(* CODESYS project i_hmi.library
   DefaultNamespace: KOSTAL.AF2024.HMI.I_Hmi
   DocFormat: reStructuredText
   Description: Base for HMI Interfaces in UTF16
   Author: Frank Dümpelmann
   Title: KOSTAL.AF2024.HMI.I_Hmi
   Version: 1.0.0.0
   Company: KOSTAL GmbH & Co.KG
   Placeholder: KOSTAL.AF2024.HMI.I_Hmi

Project tree, tasks and I/O mapping:
  libraries: KOSTAL.AF2024.Core.functionResponse, 1.0.0.0 (KOSTAL GmbH & Co.KG); KOSTAL.AF2024.Core.MainControl, 1.0.0.0 (KOSTAL GmbH & Co.KG); KOSTAL.AF2024.Core.Process, 1.0.0.0 (KOSTAL GmbH & Co.KG); KOSTAL.AF2024.Core.Settings, 1.0.0.0 (KOSTAL GmbH & Co.KG); KOSTAL.AF2024.Core.System, 1.0.0.0 (KOSTAL GmbH & Co.KG); KOSTAL.AF2024.HMI.Controls, 1.0.0.0 (KOSTAL GmbH & Co.KG)
  Aliases/
    data type T_ARTICLENAME
    data type T_BUTTON_TEXT
    data type T_F_BUTTON_TEXT
    data type T_LANGUAGENAME
    data type T_PAGE_TEXT
  DUT/
    Fn_Button/
      interface _I_T_Fn_Button: Button, clear_controls
      interface _I_T_Fn_Button_CopyFrom: CopyFrom
      interface _I_T_Fn_Button_Owner: Button_Owner, clear, clear_signals, CopyFrom
      interface _I_T_Fn_Button_RO: Button_RO, CopyTo
      data type _T_F_ButtonRange
      function block _T_Fn_Button [ST]: Button, Button_Owner, Button_RO, clear, clear_controls, clear_signals, CopyFrom, CopyTo
    Message/
      interface _I_T_Message: clear, Content, State
      interface _I_T_Message_CopyFrom: CopyFrom
      interface _I_T_Message_Owner: CopyFrom
      interface _I_T_Message_RO: Content, CopyTo, State
      function block _T_Message [ST]: clear, Content, CopyFrom, CopyTo, State
    data type E_STATE
    data type E_UserLevel
  MainControl/
    function block FB_MainControl [ST]: Button_Article_Owner, Button_Auto_Owner, Button_Door_Owner, Button_Manual_Owner, Button_OnOff_Owner, Button_Parameters_Owner, Button_Run_Owner, Button_RunEmpty_Owner, Button_Article_RO, Button_Auto_RO, Button_Door_RO, Button_Manual_RO, Button_OnOff_RO, Button_Parameters_RO, Button_Run_RO, Button_RunEmpty_RO, Button_Article, Button_Auto, Button_Door, Button_Manual, Button_OnOff, Button_Parameters, Button_RunEmpty, Button_RunStop, clear, Language, linkMainControl, Name, statusDoor_close, statusDoor_open, statusDoor_safe, UserLevel, Version_PLC
    interface I_MainControl: Button_Article, Button_Auto, Button_Door, Button_Manual, Button_OnOff, Button_Parameters, Button_RunEmpty, Button_RunStop, Language, linkMainControl, Name, statusDoor_close, statusDoor_open, statusDoor_safe, UserLevel, Version_PLC
    interface I_MainControl_Owner: Button_Article_Owner, Button_Auto_Owner, Button_Door_Owner, Button_Manual_Owner, Button_OnOff_Owner, Button_Parameters_Owner, Button_Run_Owner, Button_RunEmpty_Owner, Language, clear
    interface I_MainControl_RO: Button_Article_RO, Button_Auto_RO, Button_Door_RO, Button_Manual_RO, Button_OnOff_RO, Button_Parameters_RO, Button_Run_RO, Button_RunEmpty_RO, Language, Name, statusDoor_close, statusDoor_open, statusDoor_safe, UserLevel, Version_PLC
  Page/
    Page_Listing/
      _Buttons/
        interface _I_T_Listing_Buttons: Button_Left, Button_Right, clear_controls
        interface _I_T_Listing_Buttons_CopyFrom: CopyFrom
        interface _I_T_Listing_Buttons_Owner: Button_Left_Owner, Button_Right_Owner, clear, clear_signals, CopyFrom
        interface _I_T_Listing_Buttons_RO: Button_Right_RO, Button_RO, CopyTo
        function block _T_Listing_Buttons [ST]: Button_Left, Button_Left_Owner, Button_Right, Button_Right_Owner, Button_Right_RO, Button_RO, clear, clear_controls, clear_signals, CopyFrom, CopyTo
      _Messages/
        interface _I_T_Listing_Messages: clear, Message
        interface _I_T_Listing_Messages_CopyFrom: CopyFrom
        interface _I_T_Listing_Messages_Owner: CopyFrom, Message_Owner
        interface _I_T_Listing_Messages_RO: CopyTo, Message_RO
        function block _T_Listing_Messages [ST]: clear, CopyFrom, CopyTo, Message, Message_Owner, Message_RO
      Listing/
        function block FB_Page_Listing [ST]: Activate, Buttons, Buttons_Owner, Buttons_RO, clear, clear_buttons, clear_controls, clear_messages, clear_signals, Messages, Messages_Owner, Messages_RO
        interface I_Page_Listing: Activate, Buttons, clear_controls, clear_messages, Messages
        interface I_Page_Listing_Owner: Buttons_Owner, clear, clear_buttons, clear_signals, Messages_Owner
        interface I_Page_Listing_RO: Activate, Buttons_RO, Messages_RO
    Page_PDEF/
      _Button/
        interface _I_T_PDEF_Button_Member: State
        interface _I_T_PDEF_Button_Owner: State
        interface _I_T_PDEF_Button_RO: State
        function block _T_PDEF_Button [ST]: clear, clear_control, CopyFrom, State
      _Buttons/
        interface _I_T_PDEF_Buttons_CopyFrom: CopyFrom
        interface _I_T_PDEF_Buttons_Member: Button_Member, clear_controls
        interface _I_T_PDEF_Buttons_Owner: Button_Owner, clear, clear_signals, CopyFrom
        interface _I_T_PDEF_Buttons_RO: Button, CopyTo
        function block _T_PDEF_Buttons [ST]: Button, Button_Member, Button_Owner, clear, clear_controls, clear_signals, CopyFrom, CopyTo
      _Messages/
        interface _I_T_PDEF_Messages_CopyFrom: CopyFrom
        interface _I_T_PDEF_Messages_Member: clear, CopyFrom, Message
        interface _I_T_PDEF_Messages_Owner: Message_Owner
        interface _I_T_PDEF_Messages_RO: CopyTo, Message_RO
        function block _T_PDEF_Messages [ST]: clear, CopyFrom, CopyTo, Message, Message_Owner, Message_RO
      PDEF/
        function block FB_Page_PDEF [ST]: Buttons, Confirm, Message, Messages, Buttons_Owner, Confirm_Owner, Message_Owner, Messages_Owner, Buttons_RO, Confirm_RO, Message_RO, Messages_RO, Activate, clear, Name
        interface I_Page_PDEF: Buttons, Confirm, Message, Messages, Buttons_RO, Confirm_RO, Message_RO, Messages_RO, Activate, Name
        interface I_Page_PDEF_Owner: Buttons, Confirm, Message, Messages, Buttons_Owner, Confirm_Owner, Message_Owner, Messages_Owner, Buttons_RO, Confirm_RO, Message_RO, Messages_RO, Activate, clear, Name
        interface I_Page_PDEF_RO: Activate, Buttons_RO, Confirm_RO, Message_RO, Messages_RO, Name
    Page_Station/
      function block FB_Page_Station [ST]: Button_Enter, Button_Escape, Button_Minus, Button_OnOff, Button_Plus, Buttons_Custom, clear_controls, Name, Status, Text, Button_Enter_Owner, Button_Escape_Owner, Button_Minus_Owner, Button_OnOff_Owner, Button_Plus_Owner, Buttons_Custom_Owner, clear, clear_button, clear_signals, Status_Owner, Text_Owner, Button_Enter_RO, Button_Escape_RO, Button_Minus_RO, Button_OnOff_RO, Button_Plus_RO, Buttons_Custom_RO, Name_RO, Status_RO, Text_RO
      interface I_Page_Station: Button_Enter, Button_Escape, Button_Minus, Button_OnOff, Button_Plus, Buttons_Custom, clear_controls, Name, Status, Text
      interface I_Page_Station_Owner: Button_Enter_Owner, Button_Escape_Owner, Button_Minus_Owner, Button_OnOff_Owner, Button_Plus_Owner, Buttons_Custom_Owner, clear, clear_button, clear_signals, Status_Owner, Text_Owner
      interface I_Page_Station_RO: Button_Enter_RO, Button_Escape_RO, Button_Minus_RO, Button_OnOff_RO, Button_Plus_RO, Buttons_Custom_RO, Name, Status_RO, Text_RO
    Page_XYZ/
      _Buttons/
        interface _I_T_XYZ_Buttons: Button, clear_controls
        interface _I_T_XYZ_Buttons_CopyFrom: CopyFrom
        interface _I_T_XYZ_Buttons_Owner: Button_Owner, clear, clear_signals, CopyFrom
        interface _I_T_XYZ_Buttons_RO: Button_RO, CopyTo
        function block _T_XYZ_Buttons [ST]: Button, Button_Owner, Button_RO, clear, clear_controls, clear_signals, CopyFrom, CopyTo
      function block FB_page_XYZ [ST]: Button_Backward, Button_Down, Button_Forward, Button_Left, Button_Minus, Button_Plus, Button_Right, Button_Up, Buttons_Custom, clear_controls, SetText, Button_Backward_Owner, Button_Down_Owner, Button_Forward_Owner, Button_Left_Owner, Button_Minus_Owner, Button_Plus_Owner, Button_Right_Owner, Button_Up_Owner, Buttons_Custom_Owner, Button_Backward_RO, Button_Down_RO, Button_Forward_RO, Button_Left_RO, Button_Minus_RO, Button_Plus_RO, Button_Right_RO, Button_Up_RO, Buttons_Custom_RO, GetText, Activate, clear, clear_signals
      interface I_page_XYZ: Activate, Button_Backward, Button_Down, Button_Forward, Button_Left, Button_Minus, Button_Plus, Button_Right, Button_Up, clear_controls, SetText
      interface I_page_XYZ_Owner: Button_Backward_Owner, Button_Down_Owner, Button_Forward_Owner, Button_Left_Owner, Button_Minus_Owner, Button_Plus_Owner, Button_Right_Owner, Button_Up_Owner, clear, clear_signals
      interface I_page_XYZ_RO: Activate, Button_Backward_RO, Button_Down_RO, Button_Forward_RO, Button_Left_RO, Button_Minus_RO, Button_Plus_RO, Button_Right_RO, Button_Up_RO, GetText
  Project Information/
    function F_GetCompany [ST]
    function F_GetTitle [ST]
    function F_GetVersion [ST]
  Version/
    global variables Global_Version
  global variables GVL_CONSTANT
*)

// Aliases/T_ARTICLENAME
TYPE T_ARTICLENAME : STRING(40)
; END_TYPE

// Aliases/T_BUTTON_TEXT
TYPE T_BUTTON_TEXT : WSTRING(15)
; END_TYPE

// Aliases/T_F_BUTTON_TEXT
TYPE T_F_BUTTON_TEXT : WSTRING(10)
; END_TYPE

// Aliases/T_LANGUAGENAME
TYPE T_LANGUAGENAME : STRING(40)
; END_TYPE

// Aliases/T_PAGE_TEXT
TYPE T_PAGE_TEXT : WSTRING(255)
; END_TYPE

// DUT/Fn_Button/_T_F_ButtonRange
(*
Description
===========
| Limited data type for the index of an F-Button
*)
TYPE _T_F_ButtonRange : INT(1..8); END_TYPE

// DUT/E_STATE
(*
Description
===========
| Data type to describe a message state
*)
{attribute 'qualified_only'}
{attribute 'strict'}
TYPE E_STATE :
	(
		NONE						:=0, 
		PASS						:=1, 
		FAIL						:=2, 
		ATTENTION				:=3, 
		ERROR						:=4, 
		COMMON_REQUEST	:=5
	);
END_TYPE

// DUT/E_UserLevel
{attribute 'qualified_only'}
{attribute 'strict'}
TYPE E_UserLevel :
(
	operator := 0,
	service := 1,
	quality := 2
);
END_TYPE

// Version/Global_Version
{attribute 'TcGenerated'}
{attribute 'no-analysis'}
{attribute 'linkalways'}
// This function has been automatically generated from the project information.
VAR_GLOBAL CONSTANT
	{attribute 'const_non_replaced'}
	stLibVersion_KOSTAL_AF2024_HMI_I_Hmi : ST_LibVersion := (iMajor := 1, iMinor := 0, iBuild := 0, iRevision := 0, nFlags := 0, sVersion := '1.0.0.0');
END_VAR

// GVL_CONSTANT
{attribute 'qualified_only'}
VAR_GLOBAL CONSTANT

	MAX_FN_BUTTON	: INT:= 7;	//INT:= 7 	Maximum number of F-buttons (F8 is intern used as Help Page access)

	MAX_LISTING_LINE	: INT:= 10;	//INT:= 10	Maximum number of lines on listing page
	
	MAX_PDEF_BUTTONS	: INT:= 12;	//INT:= 12	Maximum number of FDEF buttons
	MAX_PDEF_MESSAGES	: INT:= 9;	//INT:= 9	Maximum number of FDEF messages

	MAX_XYZ_LINE	: INT:= 4;
	MAX_XYZ_BUTTON		: INT:= 4;	//INT:= 4	Maximum number of cusom Buttons on XYZ page
END_VAR

// DUT/Fn_Button/_I_T_Fn_Button
INTERFACE _I_T_Fn_Button EXTENDS _I_T_Fn_Button_RO

METHOD PUBLIC Button : KOSTAL_AF2024_HMI_Controls.I_T_Button_controlled
VAR_INPUT
	Number	: INT;
END_VAR
END_METHOD

METHOD PUBLIC clear_controls
END_METHOD

END_INTERFACE

// DUT/Fn_Button/_I_T_Fn_Button_RO
INTERFACE _I_T_Fn_Button_RO EXTENDS KOSTAL_AF2024_Core_System.I_Interface

METHOD PUBLIC Button_RO : KOSTAL_AF2024_HMI_Controls.I_T_Button_controlled
VAR_INPUT
	Number	: _T_F_ButtonRange;
END_VAR
END_METHOD

METHOD PUBLIC CopyTo
VAR_INPUT
	IN	: _I_T_Fn_Button_CopyFrom;
END_VAR
END_METHOD

END_INTERFACE

// DUT/Fn_Button/_I_T_Fn_Button_CopyFrom
INTERFACE _I_T_Fn_Button_CopyFrom EXTENDS KOSTAL_AF2024_Core_System.I_Interface

METHOD PUBLIC CopyFrom
VAR_INPUT
	IN	: _I_T_Fn_Button_RO;
END_VAR
END_METHOD

END_INTERFACE

// DUT/Fn_Button/_I_T_Fn_Button_Owner
INTERFACE _I_T_Fn_Button_Owner EXTENDS _I_T_Fn_Button

METHOD PUBLIC Button_Owner : KOSTAL_AF2024_HMI_Controls.I_T_Button_controlled_Owner
VAR_INPUT
	Number	: _T_F_ButtonRange;
END_VAR
END_METHOD

METHOD PUBLIC clear
END_METHOD

METHOD PUBLIC clear_signals
END_METHOD

METHOD PUBLIC CopyFrom
VAR_INPUT
	IN	: _I_T_Fn_Button_RO;
END_VAR
END_METHOD

END_INTERFACE

// DUT/Fn_Button/_T_Fn_Button
(*

:Author: Frank Dümpelmann <f.duempelmann@kostal.com>, Martin Hundt <m.hundt@kostal.com>
:Date: 2018-11-20

Function
========
| Data structure representing an array of buttons (FB_ControlledButton)
| Function to clear all content or signals only
*)

FUNCTION_BLOCK PUBLIC _T_Fn_Button IMPLEMENTS _I_T_Fn_Button_RO, _I_T_Fn_Button_Owner, _I_T_Fn_Button, _I_T_Fn_Button_CopyFrom

VAR
	_F		: ARRAY[1..GVL_CONSTANT.MAX_FN_BUTTON] OF KOSTAL_AF2024_HMI_Controls.T_Button_controlled;	//ARRAY[1..GVL_CONSTANT.MAX_FN_BUTTON] OF KOSTAL_TC3_Controls_button.FB_Button_controlled
	_Dummy	: KOSTAL_AF2024_HMI_Controls.T_Button_controlled;
END_VAR

METHOD PUBLIC Button : KOSTAL_AF2024_HMI_Controls.I_T_Button_controlled
VAR_INPUT
	Number	: INT;
END_VAR

IF (Number < 1) OR (Number > GVL_CONSTANT.MAX_FN_BUTTON) THEN	Button:= _Dummy;	RETURN;	END_IF

Button:= _F[Number];
END_METHOD

METHOD PUBLIC Button_Owner : KOSTAL_AF2024_HMI_Controls.I_T_Button_controlled_Owner
VAR_INPUT
	Number	: _T_F_ButtonRange;
END_VAR

IF (Number < 1) OR (Number > 8) THEN	Button_Owner:= _Dummy;	RETURN;	END_IF

Button_Owner:= _F[Number];
END_METHOD

METHOD PUBLIC Button_RO : KOSTAL_AF2024_HMI_Controls.I_T_Button_controlled
VAR_INPUT
	Number	: _T_F_ButtonRange;
END_VAR

IF (Number < 1) OR (Number > 8) THEN	Button_RO:= _Dummy;	RETURN;	END_IF

Button_RO:= _F[Number];
END_METHOD

METHOD PUBLIC clear


VAR
	_index: INT;	//INT
END_VAR

FOR _index:= 1 TO GVL_CONSTANT.MAX_FN_BUTTON DO
	_F[_index].clear();
END_FOR
END_METHOD

METHOD PUBLIC clear_controls

VAR
	_index: INT;	//INT
END_VAR

FOR _index:= 1 TO GVL_CONSTANT.MAX_FN_BUTTON DO
	_F[_index].clear_control();
END_FOR
END_METHOD

METHOD PUBLIC clear_signals

VAR
	_index: INT;	//INT
END_VAR

FOR _index:= 1 TO GVL_CONSTANT.MAX_FN_BUTTON DO
	_F[_index].clear_signals();
END_FOR
END_METHOD

METHOD PUBLIC CopyFrom
VAR_INPUT
	IN	: _I_T_Fn_Button_RO;
END_VAR

VAR
	_i: INT;
END_VAR

IF IN = 0 THEN RETURN;	END_IF

FOR _i:= 1 TO GVL_CONSTANT.MAX_FN_BUTTON DO
	_F[_i].CopyFrom(IN.Button_RO(_i));
END_FOR
END_METHOD

METHOD PUBLIC CopyTo
VAR_INPUT
	IN	: _I_T_Fn_Button_CopyFrom;
END_VAR

IF IN = 0 THEN RETURN;	END_IF

IN.CopyFrom(THIS^);
END_METHOD

END_FUNCTION_BLOCK

// DUT/Message/_I_T_Message
INTERFACE _I_T_Message EXTENDS _I_T_Message_RO

METHOD PUBLIC clear
VAR_INPUT
END_VAR
END_METHOD

PROPERTY PUBLIC Content : KOSTAL_AF2024_Core_Settings.T_MaxString
SET
END_SET
END_PROPERTY

PROPERTY PUBLIC State : E_STATE
SET
END_SET
END_PROPERTY

END_INTERFACE

// DUT/Message/_I_T_Message_RO
INTERFACE _I_T_Message_RO EXTENDS KOSTAL_AF2024_Core_System.I_Interface

PROPERTY PUBLIC Content : KOSTAL_AF2024_Core_Settings.T_MaxString
GET
END_GET
END_PROPERTY

METHOD PUBLIC CopyTo
VAR_INPUT
	IN	: _I_T_Message_CopyFrom;
END_VAR
END_METHOD

PROPERTY PUBLIC State : E_STATE
GET
END_GET
END_PROPERTY

END_INTERFACE

// DUT/Message/_I_T_Message_CopyFrom
INTERFACE _I_T_Message_CopyFrom EXTENDS KOSTAL_AF2024_Core_System.I_Interface

METHOD PUBLIC CopyFrom
VAR_INPUT
	IN	: _I_T_Message_RO;
END_VAR
END_METHOD

END_INTERFACE

// DUT/Message/_I_T_Message_Owner
INTERFACE _I_T_Message_Owner EXTENDS _I_T_Message

METHOD PUBLIC CopyFrom
VAR_INPUT
	IN	: _I_T_Message_RO;
END_VAR
END_METHOD

END_INTERFACE

// DUT/Message/_T_Message
(*

:Author: Frank Dümpelmann <f.duempelmann@kostal.com>, Martin Hundt <m.hundt@kostal.com>
:Date: 2018-11-20

Function
========
Data type representing a message with content (text) and state (error, pass,fail,...)

*)

FUNCTION_BLOCK PUBLIC _T_Message IMPLEMENTS _I_T_Message_RO, _I_T_Message_Owner, _I_T_Message, _I_T_Message_CopyFrom

VAR
	_Content	: KOSTAL_AF2024_Core_Settings.T_MaxString;
	_State		: E_STATE;
END_VAR

METHOD PUBLIC clear
VAR_INPUT
END_VAR

_Content:= "";
_State:= E_STATE.NONE;
END_METHOD

PROPERTY PUBLIC Content : KOSTAL_AF2024_Core_Settings.T_MaxString
GET

Content:= _Content;
END_GET
SET

_Content:= Content;
END_SET
END_PROPERTY

METHOD PUBLIC CopyFrom
VAR_INPUT
	IN	: _I_T_Message_RO;
END_VAR

IF IN = 0 THEN RETURN;	END_IF

_Content	:= IN.Content;
_State		:= IN.State;
END_METHOD

METHOD PUBLIC CopyTo
VAR_INPUT
	IN	: _I_T_Message_CopyFrom;
END_VAR

IF IN = 0 THEN RETURN;	END_IF

IN.CopyFrom(THIS^);
END_METHOD

PROPERTY PUBLIC State : E_STATE
GET

State:= _State;
END_GET
SET

_State:= State;
END_SET
END_PROPERTY

END_FUNCTION_BLOCK

// MainControl/FB_MainControl
(*

:Author: Frank Dümpelmann <f.duempelmann@kostal.com>, Martin Hundt <m.hundt@kostal.com>
:Date: 2020-02-20

Function
========
| Base class to implement a machine's main control

Methods and Properties
======================
| see documentation

*)
FUNCTION_BLOCK PUBLIC FB_MainControl IMPLEMENTS I_MainControl_RO, I_MainControl_Owner, I_MainControl

VAR
	_Name		: KOSTAL_AF2024_Core_Settings.T_MaxString;

	_OnOff		: KOSTAL_AF2024_HMI_Controls.T_Button_controlled;
	_RunStop	: KOSTAL_AF2024_HMI_Controls.T_Button_controlled;
	_RunEmpty	: KOSTAL_AF2024_HMI_Controls.T_Button_controlled;
                                             
	_Manual		: KOSTAL_AF2024_HMI_Controls.T_Button_controlled;
	_Auto		: KOSTAL_AF2024_HMI_Controls.T_Button_controlled;
	_Parameters		: KOSTAL_AF2024_HMI_Controls.T_Button_controlled;
	_Door		: KOSTAL_AF2024_HMI_Controls.T_Button_controlled;
	_Article	: KOSTAL_AF2024_HMI_Controls.T_Button_controlled;

	_statusDoor_close	: BOOL;	
	_statusDoor_open	: BOOL;	
	_statusDoor_safe	: BOOL;	
	
	_mainControl	: KOSTAL_AF2024_Core_MainControl.I_MainControl;

	
	_userLevel		: E_UserLevel;
	_language			: STRING;
	_version_PLC	: STRING;


END_VAR

(*
Description
===========
| Article button
*)
PROPERTY PUBLIC Button_Article_Owner : KOSTAL_AF2024_HMI_Controls.I_T_Button_controlled_Owner
GET

Button_Article_Owner := _Article;
END_GET
END_PROPERTY

(*
Description
===========
| Automatic button
*)
PROPERTY PUBLIC Button_Auto_Owner : KOSTAL_AF2024_HMI_Controls.I_T_Button_controlled_Owner
GET

Button_Auto_Owner := _Auto;
END_GET
END_PROPERTY

(*
Description
===========
| Door button
*)
PROPERTY PUBLIC Button_Door_Owner : KOSTAL_AF2024_HMI_Controls.I_T_Button_controlled_Owner
GET

Button_Door_Owner := _Door;
END_GET
END_PROPERTY

(*
Description
===========
| Manual button
*)
PROPERTY PUBLIC Button_Manual_Owner : KOSTAL_AF2024_HMI_Controls.I_T_Button_controlled_Owner
GET

Button_Manual_Owner := _Manual;
END_GET
END_PROPERTY

(*
Description
===========
| On/off button
*)
PROPERTY PUBLIC Button_OnOff_Owner : KOSTAL_AF2024_HMI_Controls.I_T_Button_controlled_Owner
GET

Button_OnOff_Owner := _OnOff;
END_GET
END_PROPERTY

(*
Description
===========
| Parameters button
*)
PROPERTY PUBLIC Button_Parameters_Owner : KOSTAL_AF2024_HMI_Controls.I_T_Button_controlled_Owner
GET

Button_Parameters_Owner := _Parameters;
END_GET
END_PROPERTY

(*
Description
===========
| Run button
*)

PROPERTY PUBLIC Button_Run_Owner : KOSTAL_AF2024_HMI_Controls.I_T_Button_controlled_Owner
GET

Button_Run_Owner := _RunStop;
END_GET
END_PROPERTY

(*
Description
===========
| Work empty button
*)
PROPERTY PUBLIC Button_RunEmpty_Owner : KOSTAL_AF2024_HMI_Controls.I_T_Button_controlled_Owner
GET

Button_RunEmpty_Owner := _RunEmpty;
END_GET
END_PROPERTY

(*
Description
===========
| Article button
*)
PROPERTY PUBLIC Button_Article_RO : KOSTAL_AF2024_HMI_Controls.I_T_Button_controlled_RO
GET
Button_Article_RO := _Article;
END_GET
END_PROPERTY

(*
Description
===========
| Automatic button
*)
PROPERTY PUBLIC Button_Auto_RO : KOSTAL_AF2024_HMI_Controls.I_T_Button_controlled_RO
GET

Button_Auto_RO := _Auto;
END_GET
END_PROPERTY

(*
Description
===========
| Door button
*)
PROPERTY PUBLIC Button_Door_RO : KOSTAL_AF2024_HMI_Controls.I_T_Button_controlled_RO
GET

Button_Door_RO := _Door;
END_GET
END_PROPERTY

(*
Description
===========
| Manual button
*)
PROPERTY PUBLIC Button_Manual_RO : KOSTAL_AF2024_HMI_Controls.I_T_Button_controlled_RO
GET

Button_Manual_RO := _Manual;
END_GET
END_PROPERTY

(*
Description
===========
| On/off button
*)
PROPERTY PUBLIC Button_OnOff_RO : KOSTAL_AF2024_HMI_Controls.I_T_Button_controlled_RO
GET

Button_OnOff_RO := _OnOff;
END_GET
END_PROPERTY

(*
Description
===========
| Parameters button
*)
PROPERTY PUBLIC Button_Parameters_RO : KOSTAL_AF2024_HMI_Controls.I_T_Button_controlled_RO
GET

Button_Parameters_RO := _Parameters;
END_GET
END_PROPERTY

(*
Description
===========
| station button
*)

PROPERTY PUBLIC Button_Run_RO : KOSTAL_AF2024_HMI_Controls.I_T_Button_controlled_RO
GET

Button_Run_RO := _RunStop;
END_GET
END_PROPERTY

(*
Description
===========
| Work empty button
*)
PROPERTY PUBLIC Button_RunEmpty_RO : KOSTAL_AF2024_HMI_Controls.I_T_Button_controlled_RO
GET

Button_RunEmpty_RO := _RunEmpty;
END_GET
END_PROPERTY

(*
Description
===========
| Article button
*)
PROPERTY PUBLIC Button_Article : KOSTAL_AF2024_HMI_Controls.I_T_Button_controlled
GET
Button_Article := _Article;
END_GET
END_PROPERTY

(*
Description
===========
| Automatic button
*)
PROPERTY PUBLIC Button_Auto : KOSTAL_AF2024_HMI_Controls.I_T_Button_controlled
GET

Button_Auto := _Auto;
END_GET
END_PROPERTY

(*
Description
===========
| Door button
*)
PROPERTY PUBLIC Button_Door : KOSTAL_AF2024_HMI_Controls.I_T_Button_controlled
GET

Button_Door := _Door;
END_GET
END_PROPERTY

(*
Description
===========
| Manual button
*)
PROPERTY PUBLIC Button_Manual : KOSTAL_AF2024_HMI_Controls.I_T_Button_controlled
GET

Button_Manual := _Manual;
END_GET
END_PROPERTY

(*
Description
===========
| On/off button
*)
PROPERTY PUBLIC Button_OnOff : KOSTAL_AF2024_HMI_Controls.I_T_Button_controlled
GET

Button_OnOff := _OnOff;
END_GET
END_PROPERTY

(*
Description
===========
| Parameters button
*)
PROPERTY PUBLIC Button_Parameters : KOSTAL_AF2024_HMI_Controls.I_T_Button_controlled
GET

Button_Parameters := _Parameters;
END_GET
END_PROPERTY

(*
Description
===========
| Work empty button
*)
PROPERTY PUBLIC Button_RunEmpty : KOSTAL_AF2024_HMI_Controls.I_T_Button_controlled
GET

Button_RunEmpty := _RunEmpty;
END_GET
END_PROPERTY

(*
Description
===========
| Run button
*)

PROPERTY PUBLIC Button_RunStop : KOSTAL_AF2024_HMI_Controls.I_T_Button_controlled
GET

Button_RunStop := _RunStop;
END_GET
END_PROPERTY

METHOD PUBLIC clear


_Name			:= "";

_OnOff.clear();
_RunStop.clear();
_RunEmpty.clear();

_Manual.clear();
_Auto.clear();
_Parameters.clear();
_Door.clear();
_Article.clear();


//_statusManual			:= FALSE;
//_statusAuto				:= FALSE;
//_statusData				:= FALSE;
_statusDoor_close	:= FALSE;
_statusDoor_open	:= FALSE;
_statusDoor_safe	:= FALSE;

//_statusOnOff			:= FALSE;
//_statusRun	:= FALSE;
//_statusWorkEmpty	:= FALSE;
END_METHOD

PROPERTY Language : STRING
GET
Language := _language;
END_GET
SET
PUBLIC 
VAR
END_VAR
_language := Language;
END_SET
END_PROPERTY

(*
Description
===========
| Link an  expert page user with index to the FlexHMI
*)
METHOD PUBLIC linkMainControl

VAR_INPUT
	control			: KOSTAL_AF2024_Core_MainControl.I_MainControl;
END_VAR

//_demand := cellDemand;
//_mode	:= cellMode;


_mainControl := control;
END_METHOD

(*
Description
===========
| Name of the machine
*)
PROPERTY PUBLIC Name : KOSTAL_AF2024_Core_Settings.T_MaxString
GET

Name:= _Name;
END_GET
SET

_Name:= Name;
END_SET
END_PROPERTY

(*
Description
===========
| Status of the door(s) is closed
*)
PROPERTY PUBLIC statusDoor_close : BOOL
GET

statusDoor_close:= _statusDoor_close;
END_GET
SET

_statusDoor_close:= statusDoor_close;
END_SET
END_PROPERTY

(*
Description
===========
| Status of the door(s) is open
*)
PROPERTY PUBLIC statusDoor_open : BOOL
GET

statusDoor_open:= _statusDoor_open;
END_GET
SET

_statusDoor_open:= statusDoor_open;
END_SET
END_PROPERTY

(*
Description
===========
| Status of the door(s) is safe (closed and locked)
*)
PROPERTY PUBLIC statusDoor_safe : BOOL
GET

statusDoor_safe:= _statusDoor_safe;
END_GET
SET

_statusDoor_safe:= statusDoor_safe;
END_SET
END_PROPERTY

PROPERTY PUBLIC UserLevel : E_UserLevel
GET
UserLevel := _userLevel;
END_GET
SET
_userLevel := UserLevel;
END_SET
END_PROPERTY

PROPERTY Version_PLC : String
GET
Version_PLC := _version_PLC;
END_GET
SET
_version_PLC := Version_PLC;
END_SET
END_PROPERTY

END_FUNCTION_BLOCK

// MainControl/I_MainControl_RO
INTERFACE I_MainControl_RO EXTENDS KOSTAL_AF2024_Core_System.I_Interface

(*
Description
===========
| Article button
*)
PROPERTY PUBLIC Button_Article_RO : KOSTAL_AF2024_HMI_Controls.I_T_Button_controlled_RO
GET
END_GET
END_PROPERTY

(*
Description
===========
| Automatic button
*)
PROPERTY PUBLIC Button_Auto_RO : KOSTAL_AF2024_HMI_Controls.I_T_Button_controlled_RO
GET
END_GET
END_PROPERTY

(*
Description
===========
| Door button
*)
PROPERTY PUBLIC Button_Door_RO : KOSTAL_AF2024_HMI_Controls.I_T_Button_controlled_RO
GET
END_GET
END_PROPERTY

(*
Description
===========
| Manual button
*)
PROPERTY PUBLIC Button_Manual_RO : KOSTAL_AF2024_HMI_Controls.I_T_Button_controlled_RO
GET
END_GET
END_PROPERTY

(*
Description
===========
| On/off button
*)
PROPERTY PUBLIC Button_OnOff_RO : KOSTAL_AF2024_HMI_Controls.I_T_Button_controlled_RO
GET
END_GET
END_PROPERTY

(*
Description
===========
| Parameters button
*)
PROPERTY PUBLIC Button_Parameters_RO : KOSTAL_AF2024_HMI_Controls.I_T_Button_controlled_RO
GET
END_GET
END_PROPERTY

(*
Description
===========
| Run button
*)

PROPERTY PUBLIC Button_Run_RO : KOSTAL_AF2024_HMI_Controls.I_T_Button_controlled_RO
GET
END_GET
END_PROPERTY

(*
Description
===========
| Work empty button
*)
PROPERTY PUBLIC Button_RunEmpty_RO : KOSTAL_AF2024_HMI_Controls.I_T_Button_controlled_RO
GET
END_GET
END_PROPERTY

PROPERTY Language : STRING
GET
END_GET
END_PROPERTY

PROPERTY PUBLIC Name : KOSTAL_AF2024_Core_Settings.T_MaxString
GET
END_GET
END_PROPERTY

PROPERTY PUBLIC statusDoor_close : BOOL
GET
END_GET
END_PROPERTY

PROPERTY PUBLIC statusDoor_open : BOOL
GET
END_GET
END_PROPERTY

PROPERTY PUBLIC statusDoor_safe : BOOL
GET
END_GET
END_PROPERTY

PROPERTY PUBLIC UserLevel : E_UserLevel
GET
END_GET
END_PROPERTY

PROPERTY Version_PLC : String
GET
END_GET
END_PROPERTY

END_INTERFACE

// MainControl/I_MainControl_Owner
INTERFACE I_MainControl_Owner EXTENDS I_MainControl

(*
Description
===========
| Article button
*)
PROPERTY PUBLIC Button_Article_Owner : KOSTAL_AF2024_HMI_Controls.I_T_Button_controlled_Owner
GET
END_GET
END_PROPERTY

(*
Description
===========
| Automatic button
*)
PROPERTY PUBLIC Button_Auto_Owner : KOSTAL_AF2024_HMI_Controls.I_T_Button_controlled_Owner
GET
END_GET
END_PROPERTY

(*
Description
===========
| Door button
*)
PROPERTY PUBLIC Button_Door_Owner : KOSTAL_AF2024_HMI_Controls.I_T_Button_controlled_Owner
GET
END_GET
END_PROPERTY

(*
Description
===========
| Manual button
*)
PROPERTY PUBLIC Button_Manual_Owner : KOSTAL_AF2024_HMI_Controls.I_T_Button_controlled_Owner
GET
END_GET
END_PROPERTY

(*
Description
===========
| On/off button
*)
PROPERTY PUBLIC Button_OnOff_Owner : KOSTAL_AF2024_HMI_Controls.I_T_Button_controlled_Owner
GET
END_GET
END_PROPERTY

(*
Description
===========
| Parameters button
*)
PROPERTY PUBLIC Button_Parameters_Owner : KOSTAL_AF2024_HMI_Controls.I_T_Button_controlled_Owner
GET
END_GET
END_PROPERTY

(*
Description
===========
| Run button
*)

PROPERTY PUBLIC Button_Run_Owner : KOSTAL_AF2024_HMI_Controls.I_T_Button_controlled_Owner
GET
END_GET
END_PROPERTY

(*
Description
===========
| Work empty button
*)
PROPERTY PUBLIC Button_RunEmpty_Owner : KOSTAL_AF2024_HMI_Controls.I_T_Button_controlled_Owner
GET
END_GET
END_PROPERTY

PROPERTY Language : STRING
GET
END_GET
END_PROPERTY

METHOD PUBLIC clear
END_METHOD

END_INTERFACE

// MainControl/I_MainControl
INTERFACE I_MainControl EXTENDS I_MainControl_RO

(*
Description
===========
| Article button
*)
PROPERTY PUBLIC Button_Article : KOSTAL_AF2024_HMI_Controls.I_T_Button_controlled
GET
END_GET
END_PROPERTY

(*
Description
===========
| Automatic button
*)
PROPERTY PUBLIC Button_Auto : KOSTAL_AF2024_HMI_Controls.I_T_Button_controlled
GET
END_GET
END_PROPERTY

(*
Description
===========
| Door button
*)
PROPERTY PUBLIC Button_Door : KOSTAL_AF2024_HMI_Controls.I_T_Button_controlled
GET
END_GET
END_PROPERTY

(*
Description
===========
| Manual button
*)
PROPERTY PUBLIC Button_Manual : KOSTAL_AF2024_HMI_Controls.I_T_Button_controlled
GET
END_GET
END_PROPERTY

(*
Description
===========
| On/off button
*)
PROPERTY PUBLIC Button_OnOff : KOSTAL_AF2024_HMI_Controls.I_T_Button_controlled
GET
END_GET
END_PROPERTY

(*
Description
===========
| Parameters button
*)
PROPERTY PUBLIC Button_Parameters : KOSTAL_AF2024_HMI_Controls.I_T_Button_controlled
GET
END_GET
END_PROPERTY

(*
Description
===========
| Work empty button
*)
PROPERTY PUBLIC Button_RunEmpty : KOSTAL_AF2024_HMI_Controls.I_T_Button_controlled
GET
END_GET
END_PROPERTY

(*
Description
===========
| Run button
*)

PROPERTY PUBLIC Button_RunStop : KOSTAL_AF2024_HMI_Controls.I_T_Button_controlled
GET
END_GET
END_PROPERTY

PROPERTY Language : STRING
GET
END_GET
END_PROPERTY

(*
Description
===========
| Link an  expert page user with index to the FlexHMI
*)
METHOD PUBLIC linkMainControl

VAR_INPUT
	control			: KOSTAL_AF2024_Core_MainControl.I_MainControl;
END_VAR
END_METHOD

PROPERTY PUBLIC Name : KOSTAL_AF2024_Core_Settings.T_MaxString
SET
END_SET
END_PROPERTY

PROPERTY PUBLIC statusDoor_close : BOOL
SET
END_SET
END_PROPERTY

PROPERTY PUBLIC statusDoor_open : BOOL
SET
END_SET
END_PROPERTY

PROPERTY PUBLIC statusDoor_safe : BOOL
SET
END_SET
END_PROPERTY

PROPERTY PUBLIC UserLevel : E_UserLevel
SET
END_SET
END_PROPERTY

PROPERTY Version_PLC : String
SET
END_SET
END_PROPERTY

END_INTERFACE

// Page/Page_Listing/_Buttons/_I_T_Listing_Buttons
INTERFACE _I_T_Listing_Buttons EXTENDS _I_T_Listing_Buttons_RO

METHOD PUBLIC Button_Left : KOSTAL_AF2024_HMI_Controls.I_T_Button_controlled
VAR_INPUT
	Number	: INT;
END_VAR
END_METHOD

METHOD PUBLIC Button_Right : KOSTAL_AF2024_HMI_Controls.I_T_Button_controlled
VAR_INPUT
	Number	: INT;
END_VAR
END_METHOD

METHOD PUBLIC clear_controls
END_METHOD

END_INTERFACE

// Page/Page_Listing/_Buttons/_I_T_Listing_Buttons_RO
INTERFACE _I_T_Listing_Buttons_RO EXTENDS KOSTAL_AF2024_Core_System.I_Interface

METHOD PUBLIC Button_Right_RO : KOSTAL_AF2024_HMI_Controls.I_T_Button_controlled_RO
VAR_INPUT
	Number	: INT;
END_VAR
END_METHOD

METHOD PUBLIC Button_RO : KOSTAL_AF2024_HMI_Controls.I_T_Button_controlled_RO
VAR_INPUT
	Number	: INT;
END_VAR
END_METHOD

METHOD PUBLIC CopyTo
VAR_INPUT
END_VAR
END_METHOD

END_INTERFACE

// Page/Page_Listing/_Buttons/_I_T_Listing_Buttons_CopyFrom
INTERFACE _I_T_Listing_Buttons_CopyFrom EXTENDS KOSTAL_AF2024_Core_System.I_Interface

METHOD PUBLIC CopyFrom
VAR_INPUT
	IN	: _I_T_Listing_Buttons_RO;
END_VAR
END_METHOD

END_INTERFACE

// Page/Page_Listing/_Buttons/_I_T_Listing_Buttons_Owner
INTERFACE _I_T_Listing_Buttons_Owner EXTENDS _I_T_Listing_Buttons

METHOD PUBLIC Button_Left_Owner : KOSTAL_AF2024_HMI_Controls.I_T_Button_controlled_Owner
VAR_INPUT
	Number	: INT;
END_VAR
END_METHOD

METHOD PUBLIC Button_Right_Owner : KOSTAL_AF2024_HMI_Controls.I_T_Button_controlled_Owner
VAR_INPUT
	Number	: INT;
END_VAR
END_METHOD

METHOD PUBLIC clear
END_METHOD

METHOD PUBLIC clear_signals
END_METHOD

METHOD PUBLIC CopyFrom
VAR_INPUT
	IN	: _I_T_Listing_Buttons_RO;
END_VAR
END_METHOD

END_INTERFACE

// Page/Page_Listing/_Buttons/_T_Listing_Buttons
(*

:Author: Frank Dümpelmann <f.duempelmann@kostal.com>, Martin Hundt <m.hundt@kostal.com>
:Date: 2018-11-20

Function
========
Data structure representing the buttons in the listing page of the user interface

Methods and Properties
======================
| Left: Array with Buttons on the left side of the page (see FB_Button_controlled)
| Right: Array with Buttons on the right side of the page (see FB_Button_controlled)
| clear signals of buttons
| clear all buttons
*)
FUNCTION_BLOCK _T_Listing_Buttons IMPLEMENTS _I_T_Listing_Buttons_RO, _I_T_Listing_Buttons_Owner, _I_T_Listing_Buttons, _I_T_Listing_Buttons_CopyFrom

VAR
	_Left	: ARRAY[1..GVL_CONSTANT.MAX_LISTING_LINE] OF KOSTAL_AF2024_HMI_Controls.T_Button_controlled;
	_Right	: ARRAY[1..GVL_CONSTANT.MAX_LISTING_LINE] OF KOSTAL_AF2024_HMI_Controls.T_Button_controlled;

	_Dummy	: KOSTAL_AF2024_HMI_Controls.T_Button_controlled;
END_VAR

METHOD PUBLIC Button_Left : KOSTAL_AF2024_HMI_Controls.I_T_Button_controlled
VAR_INPUT
	Number	: INT;
END_VAR

IF (Number < 1) OR (Number > GVL_CONSTANT.MAX_LISTING_LINE) THEN	
	Button_Left:= _Dummy;	
	RETURN;	
END_IF

	
Button_Left:= _Left[Number];
END_METHOD

METHOD PUBLIC Button_Left_Owner : KOSTAL_AF2024_HMI_Controls.I_T_Button_controlled_Owner
VAR_INPUT
	Number	: INT;
END_VAR

IF (Number < 1) OR (Number > GVL_CONSTANT.MAX_LISTING_LINE) THEN	
	Button_Left_Owner:= _Dummy;	
	RETURN;	
END_IF

	
Button_Left_Owner:= _Left[Number];
END_METHOD

METHOD PUBLIC Button_Right : KOSTAL_AF2024_HMI_Controls.I_T_Button_controlled
VAR_INPUT
	Number	: INT;
END_VAR

IF (Number < 1) OR (Number > GVL_CONSTANT.MAX_LISTING_LINE) THEN	
	Button_Right:= _Dummy;	
	RETURN;	
END_IF

	
Button_Right:= _Right[Number];
END_METHOD

METHOD PUBLIC Button_Right_Owner : KOSTAL_AF2024_HMI_Controls.I_T_Button_controlled_Owner
VAR_INPUT
	Number	: INT;
END_VAR

IF (Number < 1) OR (Number > GVL_CONSTANT.MAX_LISTING_LINE) THEN	
	Button_Right_Owner:= _Dummy;	
	RETURN;	
END_IF

	
Button_Right_Owner:= _Right[Number];
END_METHOD

METHOD PUBLIC Button_Right_RO : KOSTAL_AF2024_HMI_Controls.I_T_Button_controlled_RO
VAR_INPUT
	Number	: INT;
END_VAR

IF (Number < 1) OR (Number > GVL_CONSTANT.MAX_LISTING_LINE) THEN	
	Button_Right_RO:= _Dummy;	
	RETURN;	
END_IF

	
Button_Right_RO:= _Right[Number];
END_METHOD

METHOD PUBLIC Button_RO : KOSTAL_AF2024_HMI_Controls.I_T_Button_controlled_RO
VAR_INPUT
	Number	: INT;
END_VAR

IF (Number < 1) OR (Number > GVL_CONSTANT.MAX_LISTING_LINE) THEN	
	Button_RO:= _Dummy;	
	RETURN;	
END_IF

	
Button_RO:= _Left[Number];
END_METHOD

METHOD PUBLIC clear


VAR
	_index: INT;	//INT
END_VAR


FOR _index:= 1 TO GVL_CONSTANT.MAX_LISTING_LINE DO
	_Left[_index].clear();
	_Right[_index].clear();
END_FOR
END_METHOD

METHOD PUBLIC clear_controls


VAR
	_index: INT;	//INT
END_VAR


FOR _index:= 1 TO GVL_CONSTANT.MAX_LISTING_LINE DO
	_Left[_index].clear_control();
	_Right[_index].clear_control();
END_FOR
END_METHOD

METHOD PUBLIC clear_signals


VAR
	_index: INT;	//INT
END_VAR


FOR _index:= 1 TO GVL_CONSTANT.MAX_LISTING_LINE DO
	_Left[_index].clear_signals();
	_Right[_index].clear_signals();
END_FOR
END_METHOD

METHOD PUBLIC CopyFrom
VAR_INPUT
	IN	: _I_T_Listing_Buttons_RO;
END_VAR

VAR
	_i: INT;
END_VAR

IF IN = 0 THEN RETURN;	END_IF

FOR _i:= 1 TO GVL_CONSTANT.MAX_LISTING_LINE DO
	_Left[_i].CopyFrom(IN.Button_RO(_i));
	_Right[_i].CopyFrom(IN.Button_Right_RO(_i));
END_FOR
END_METHOD

METHOD PUBLIC CopyTo
VAR_INPUT
END_VAR
END_METHOD

END_FUNCTION_BLOCK

// Page/Page_Listing/_Messages/_I_T_Listing_Messages
INTERFACE _I_T_Listing_Messages EXTENDS _I_T_Listing_Messages_RO

METHOD PUBLIC clear
END_METHOD

METHOD PUBLIC Message : _I_T_Message
VAR_INPUT
	Line	: INT;
END_VAR
END_METHOD

END_INTERFACE

// Page/Page_Listing/_Messages/_I_T_Listing_Messages_RO
INTERFACE _I_T_Listing_Messages_RO EXTENDS KOSTAL_AF2024_Core_System.I_Interface

METHOD PUBLIC CopyTo
VAR_INPUT
	IN	: _I_T_Listing_Messages_CopyFrom;
END_VAR
END_METHOD

METHOD PUBLIC Message_RO : _I_T_Message_RO
VAR_INPUT
	Line	: INT;
END_VAR
END_METHOD

END_INTERFACE

// Page/Page_Listing/_Messages/_I_T_Listing_Messages_CopyFrom
INTERFACE _I_T_Listing_Messages_CopyFrom EXTENDS KOSTAL_AF2024_Core_System.I_Interface

METHOD PUBLIC CopyFrom
VAR_INPUT
	IN	: _I_T_Listing_Messages_RO;
END_VAR
END_METHOD

END_INTERFACE

// Page/Page_Listing/_Messages/_I_T_Listing_Messages_Owner
INTERFACE _I_T_Listing_Messages_Owner EXTENDS _I_T_Listing_Messages

METHOD PUBLIC CopyFrom
VAR_INPUT
	IN	: _I_T_Listing_Messages_RO;
END_VAR
END_METHOD

METHOD PUBLIC Message_Owner : _I_T_Message_Owner
VAR_INPUT
	Line		: INT;
	Message	: _I_T_Message_RO;	
END_VAR
END_METHOD

END_INTERFACE

// Page/Page_Listing/_Messages/_T_Listing_Messages
(*
:Author: Frank Dümpelmann <f.duempelmann@kostal.com>, Martin Hundt <m.hundt@kostal.com>
:Date: 2018-11-20

Function
========
Data structure representing the messages in the listing page of the user interface

Methods and Properties
======================
| Line: Array of FB_Message 
| Clear: clear all messages
*)
FUNCTION_BLOCK _T_Listing_Messages IMPLEMENTS _I_T_Listing_Messages_RO, _I_T_Listing_Messages_Owner, _I_T_Listing_Messages, _I_T_Listing_Messages_CopyFrom

VAR
	_Line	:	ARRAY[1..GVL_CONSTANT.MAX_LISTING_LINE] OF _T_Message;	//ARRAY[1..GVL.LISTING_MAX_LINE] OF FB_Message
	_Dummy	: _T_Message;
END_VAR

METHOD PUBLIC clear


VAR
	_index: INT;	//INT
END_VAR




FOR _index:= 1 TO GVL_CONSTANT.MAX_LISTING_LINE DO
	_Line[_index].clear();
END_FOR
END_METHOD

METHOD PUBLIC CopyFrom
VAR_INPUT
	IN	: _I_T_Listing_Messages_RO;
END_VAR

VAR
	_i: INT;
END_VAR

IF IN = 0 THEN RETURN;	END_IF

FOR _i:= 1 TO GVL_CONSTANT.MAX_LISTING_LINE DO
	_Line[_i].CopyFrom(IN.Message_RO(INT_TO_USINT(_i)));
END_FOR
END_METHOD

METHOD PUBLIC CopyTo
VAR_INPUT
	IN	: _I_T_Listing_Messages_CopyFrom;
END_VAR

IF IN = 0 THEN RETURN;	END_IF

IN.CopyFrom(THIS^);
END_METHOD

METHOD PUBLIC Message : _I_T_Message
VAR_INPUT
	Line	: INT;
END_VAR
IF (Line < 1) OR (Line > GVL_CONSTANT.MAX_LISTING_LINE) THEN Message:= _Dummy;	RETURN;	END_IF

Message:= _Line[Line];
END_METHOD

METHOD PUBLIC Message_Owner : _I_T_Message_Owner
VAR_INPUT
	Line	: INT;
	Message	: _I_T_Message_RO;	
END_VAR
IF (Line < 1) OR (Line > GVL_CONSTANT.MAX_LISTING_LINE) THEN Message_Owner:= _Dummy;	RETURN;	END_IF

IF Message <> 0 THEN _Line[Line].CopyFrom(Message);	END_IF

Message_Owner:= _Line[Line];
END_METHOD

METHOD PUBLIC Message_RO : _I_T_Message_RO
VAR_INPUT
	Line	: INT;
END_VAR
IF (Line < 1) OR (Line > GVL_CONSTANT.MAX_LISTING_LINE) THEN Message_RO:= _Dummy;	RETURN;	END_IF

Message_RO:= _Line[Line];
END_METHOD

END_FUNCTION_BLOCK

// Page/Page_Listing/Listing/FB_Page_Listing
(*
:Author: Frank Dümpelmann <f.duempelmann@kostal.com>, Martin Hundt <m.hundt@kostal.com>
:Date: 2018-11-20

Function
========
Data structure representing the listing page in the user interface

Methods and Properties
======================
| Activate: Activate the Form
| Deactivate: Deactivate the Form
| IsActiv: Response the state of the Form
| Buttons: see FB_LISTING_Buttons
| Messages: see FB_LISTING_Messages
*)
FUNCTION_BLOCK FB_Page_Listing IMPLEMENTS I_Page_Listing_RO, I_Page_Listing_Owner, I_Page_Listing

VAR
	_Activate		: BOOL;	//BOOL	-	Activate the Form
	_Deactivate		: BOOL;	//BOOL	-	Deactivate the Form
	_IsActiv		: BOOL;	//BOOL	-	Response the state of the Form

	_Buttons	: _T_Listing_Buttons;	//FB_LISTING_Buttons
	_Messages	: _T_Listing_Messages;	//FB_LISTING_Messages
END_VAR

PROPERTY PUBLIC Activate : BOOL
GET

Activate:= _Activate;
END_GET
SET

_Activate:= Activate;
END_SET
END_PROPERTY

PROPERTY PUBLIC Buttons : _I_T_Listing_Buttons
GET

Buttons := _Buttons;
END_GET
END_PROPERTY

PROPERTY PUBLIC Buttons_Owner : _I_T_Listing_Buttons_Owner
GET

Buttons_Owner := _Buttons;
END_GET
END_PROPERTY

PROPERTY PUBLIC Buttons_RO : _I_T_Listing_Buttons_RO
GET

Buttons_RO := _Buttons;
END_GET
END_PROPERTY

METHOD PUBLIC clear


_Activate		:= FALSE;
_Deactivate	:= FALSE;
_IsActiv		:= FALSE;


_Buttons.clear();
_Messages.clear();
END_METHOD

METHOD PUBLIC clear_buttons


_Buttons.clear();
END_METHOD

METHOD PUBLIC clear_controls


_Buttons.clear_controls();
END_METHOD

METHOD PUBLIC clear_messages


_Messages.clear();
END_METHOD

METHOD PUBLIC clear_signals


_Buttons.clear_signals();
END_METHOD

PROPERTY PUBLIC Messages : _I_T_Listing_Messages
GET

Messages := _Messages;
END_GET
END_PROPERTY

PROPERTY PUBLIC Messages_Owner : _I_T_Listing_Messages_Owner
GET

Messages_Owner := _Messages;
END_GET
END_PROPERTY

PROPERTY PUBLIC Messages_RO : _I_T_Listing_Messages_RO
GET

Messages_RO := _Messages;
END_GET
END_PROPERTY

END_FUNCTION_BLOCK

// Page/Page_Listing/Listing/I_Page_Listing_RO
INTERFACE I_Page_Listing_RO EXTENDS KOSTAL_AF2024_Core_System.I_Interface

PROPERTY PUBLIC Activate : BOOL
GET
END_GET
END_PROPERTY

PROPERTY PUBLIC Buttons_RO : _I_T_Listing_Buttons_RO
GET
END_GET
END_PROPERTY

PROPERTY PUBLIC Messages_RO : _I_T_Listing_Messages_RO
GET
END_GET
END_PROPERTY

END_INTERFACE

// Page/Page_Listing/Listing/I_Page_Listing_Owner
INTERFACE I_Page_Listing_Owner EXTENDS I_Page_Listing

PROPERTY PUBLIC Buttons_Owner : _I_T_Listing_Buttons_Owner
GET
END_GET
END_PROPERTY

METHOD PUBLIC clear
END_METHOD

METHOD PUBLIC clear_buttons
END_METHOD

METHOD PUBLIC clear_signals
END_METHOD

PROPERTY PUBLIC Messages_Owner : _I_T_Listing_Messages_Owner
GET
END_GET
END_PROPERTY

END_INTERFACE

// Page/Page_Listing/Listing/I_Page_Listing
INTERFACE I_Page_Listing EXTENDS I_Page_Listing_RO

PROPERTY PUBLIC Activate : BOOL
SET
END_SET
END_PROPERTY

PROPERTY PUBLIC Buttons : _I_T_Listing_Buttons
GET
END_GET
END_PROPERTY

METHOD PUBLIC clear_controls
END_METHOD

METHOD PUBLIC clear_messages
END_METHOD

PROPERTY PUBLIC Messages : _I_T_Listing_Messages
GET
END_GET
END_PROPERTY

END_INTERFACE

// Page/Page_PDEF/_Button/_I_T_PDEF_Button_Member
INTERFACE _I_T_PDEF_Button_Member EXTENDS KOSTAL_AF2024_HMI_Controls.I_T_Button_controlled

PROPERTY PUBLIC State : E_STATE
GET
END_GET
SET
END_SET
END_PROPERTY

END_INTERFACE

// Page/Page_PDEF/_Button/_I_T_PDEF_Button_Owner
INTERFACE _I_T_PDEF_Button_Owner EXTENDS KOSTAL_AF2024_HMI_Controls.I_T_Button_controlled_Owner

PROPERTY PUBLIC State : E_STATE
GET
END_GET
SET
END_SET
END_PROPERTY

END_INTERFACE

// Page/Page_PDEF/_Button/_I_T_PDEF_Button_RO
INTERFACE _I_T_PDEF_Button_RO EXTENDS KOSTAL_AF2024_HMI_Controls.I_T_Button_controlled

PROPERTY PUBLIC State : E_STATE
GET
END_GET
END_PROPERTY

END_INTERFACE

// Page/Page_PDEF/_Button/_T_PDEF_Button
(*
Description
===========
| Extension of FB_Button_controlled with an additional state
| See documentation of FB_Button_controlled and E_STATE
*)
FUNCTION_BLOCK _T_PDEF_Button EXTENDS KOSTAL_AF2024_HMI_Controls.T_Button_controlled IMPLEMENTS _I_T_PDEF_Button_RO, _I_T_PDEF_Button_Owner, _I_T_PDEF_Button_Member

VAR
	_State	:	E_STATE;	//E_STATE
END_VAR

METHOD PUBLIC clear

_State:= E_STATE.NONE;

SUPER^.clear();
END_METHOD

METHOD PUBLIC clear_control

_State:= E_STATE.NONE;

SUPER^.clear_control();
END_METHOD

METHOD PUBLIC CopyFrom
VAR_INPUT
	IN	: KOSTAL_AF2024_HMI_Controls.I_T_Button;
END_VAR

VAR
	_oPDEF	: _I_T_PDEF_Button_RO;
END_VAR

IF IN = 0 THEN RETURN;	END_IF

IF NOT __QUERYINTERFACE(IN, _oPDEF) THEN RETURN; END_IF
IF _oPDEF = 0 THEN RETURN;	END_IF

_State:= _oPDEF.State;

SUPER^.CopyFrom(IN);
END_METHOD

PROPERTY PUBLIC State : E_STATE
GET

State:= _State;
END_GET
SET

_State:= State;
END_SET
END_PROPERTY

END_FUNCTION_BLOCK

// Page/Page_PDEF/_Buttons/_I_T_PDEF_Buttons_CopyFrom
INTERFACE _I_T_PDEF_Buttons_CopyFrom EXTENDS KOSTAL_AF2024_Core_System.I_Interface

METHOD PUBLIC CopyFrom
VAR_INPUT
	IN	: _I_T_PDEF_Buttons_RO;
END_VAR
END_METHOD

END_INTERFACE

// Page/Page_PDEF/_Buttons/_I_T_PDEF_Buttons_RO
INTERFACE _I_T_PDEF_Buttons_RO EXTENDS KOSTAL_AF2024_Core_System.I_Interface

METHOD PUBLIC Button : _I_T_PDEF_Button_RO
VAR_INPUT
	Number	: INT;
END_VAR
END_METHOD

METHOD PUBLIC CopyTo
VAR_INPUT
	IN	: _I_T_PDEF_Buttons_CopyFrom;
END_VAR
END_METHOD

END_INTERFACE

// Page/Page_PDEF/_Buttons/_I_T_PDEF_Buttons_Member
INTERFACE _I_T_PDEF_Buttons_Member EXTENDS _I_T_PDEF_Buttons_RO

METHOD PUBLIC Button_Member : _I_T_PDEF_Button_Member
VAR_INPUT
	Number	: INT;
END_VAR
END_METHOD

METHOD PUBLIC clear_controls
VAR_INPUT
END_VAR
END_METHOD

END_INTERFACE

// Page/Page_PDEF/_Buttons/_I_T_PDEF_Buttons_Owner
INTERFACE _I_T_PDEF_Buttons_Owner EXTENDS _I_T_PDEF_Buttons_Member

METHOD PUBLIC Button_Owner : _I_T_PDEF_Button_Owner
VAR_INPUT
	Number	: INT;
END_VAR
END_METHOD

METHOD PUBLIC clear
VAR_INPUT
END_VAR
END_METHOD

METHOD PUBLIC clear_signals
VAR_INPUT
END_VAR
END_METHOD

METHOD PUBLIC CopyFrom
VAR_INPUT
	IN	: _I_T_PDEF_Buttons_RO;
END_VAR
END_METHOD

END_INTERFACE

// Page/Page_PDEF/_Buttons/_T_PDEF_Buttons
(*
Description
===========
| Index: Array of buttons on the PDEF page
| Methods to clear signals or clear all
*)
FUNCTION_BLOCK PUBLIC _T_PDEF_Buttons IMPLEMENTS _I_T_PDEF_Buttons_RO, _I_T_PDEF_Buttons_Owner, _I_T_PDEF_Buttons_Member, _I_T_PDEF_Buttons_CopyFrom

VAR
	_Index	: ARRAY[1..GVL_CONSTANT.MAX_PDEF_BUTTONS] OF _T_PDEF_Button;	//ARRAY[1..GVL.MAX_PDEF_BUTTONS] OF FB_PDEF_Button
	_Dummy	: _T_PDEF_Button;
END_VAR

METHOD PUBLIC Button : _I_T_PDEF_Button_RO
VAR_INPUT
	Number	: INT;
END_VAR

IF (Number < 1) OR (Number > GVL_CONSTANT.MAX_PDEF_BUTTONS) THEN	Button:= _Dummy;	RETURN;	END_IF

Button:= _Index[Number];
END_METHOD

METHOD PUBLIC Button_Member : _I_T_PDEF_Button_Member
VAR_INPUT
	Number	: INT;
END_VAR

IF (Number < 1) OR (Number > GVL_CONSTANT.MAX_PDEF_BUTTONS) THEN	Button_Member:= _Dummy;	RETURN;	END_IF

Button_Member:= _Index[Number];
END_METHOD

METHOD PUBLIC Button_Owner : _I_T_PDEF_Button_Owner
VAR_INPUT
	Number	: INT;
END_VAR

IF (Number < 1) OR (Number > GVL_CONSTANT.MAX_PDEF_BUTTONS) THEN	Button_Owner:= _Dummy;	RETURN;	END_IF

//IF Button <> 0 THEN	_Index[Number].CopyFrom(Button);	END_IF

Button_Owner:= _Index[Number];
END_METHOD

METHOD PUBLIC clear
VAR_INPUT
END_VAR

VAR
	_i: INT;	//INT
END_VAR


FOR _i:= 1 TO GVL_CONSTANT.MAX_PDEF_BUTTONS DO
		_Index[_i].clear();
END_FOR
END_METHOD

METHOD PUBLIC clear_controls
VAR_INPUT
END_VAR

VAR
	_i: INT;	//INT
END_VAR


FOR _i:= 1 TO GVL_CONSTANT.MAX_PDEF_BUTTONS DO
	_Index[_i].clear_control();
END_FOR
END_METHOD

METHOD PUBLIC clear_signals
VAR_INPUT
END_VAR

VAR
	_i: INT;	//INT
END_VAR


FOR _i:= 1 TO GVL_CONSTANT.MAX_PDEF_BUTTONS DO
	_Index[_i].clear_signals();
END_FOR
END_METHOD

METHOD PUBLIC CopyFrom
VAR_INPUT
	IN	: _I_T_PDEF_Buttons_RO;
END_VAR

VAR
	_i: INT;
END_VAR

IF IN = 0 THEN RETURN;	END_IF

FOR _i:= 1 TO GVL_CONSTANT.MAX_PDEF_BUTTONS DO
	_Index[_i].CopyFrom(IN.Button(_i));
END_FOR
END_METHOD

METHOD PUBLIC CopyTo
VAR_INPUT
	IN	: _I_T_PDEF_Buttons_CopyFrom;
END_VAR

IF IN = 0 THEN RETURN;	END_IF

IN.CopyFrom(THIS^);
END_METHOD

END_FUNCTION_BLOCK

// Page/Page_PDEF/_Messages/_I_T_PDEF_Messages_CopyFrom
INTERFACE _I_T_PDEF_Messages_CopyFrom EXTENDS KOSTAL_AF2024_Core_System.I_Interface

METHOD PUBLIC CopyFrom
VAR_INPUT
	IN	: _I_T_PDEF_Messages_RO;
END_VAR
END_METHOD

END_INTERFACE

// Page/Page_PDEF/_Messages/_I_T_PDEF_Messages_RO
INTERFACE _I_T_PDEF_Messages_RO EXTENDS KOSTAL_AF2024_Core_System.I_Interface

METHOD PUBLIC CopyTo
VAR_INPUT
	IN	: _I_T_PDEF_Messages_CopyFrom;
END_VAR
END_METHOD

METHOD PUBLIC Message_RO : _I_T_Message_RO
VAR_INPUT
	Number	: INT;
END_VAR
END_METHOD

END_INTERFACE

// Page/Page_PDEF/_Messages/_I_T_PDEF_Messages_Member
INTERFACE _I_T_PDEF_Messages_Member EXTENDS _I_T_PDEF_Messages_RO

METHOD PUBLIC clear
END_METHOD

METHOD PUBLIC CopyFrom
VAR_INPUT
	IN	: _I_T_PDEF_Messages_RO;
END_VAR
END_METHOD

METHOD PUBLIC Message : _I_T_Message
VAR_INPUT
	Number	: INT;
END_VAR
END_METHOD

END_INTERFACE

// Page/Page_PDEF/_Messages/_I_T_PDEF_Messages_Owner
INTERFACE _I_T_PDEF_Messages_Owner EXTENDS _I_T_PDEF_Messages_Member

METHOD PUBLIC Message_Owner : _I_T_Message_Owner
VAR_INPUT
	Number	: INT;
END_VAR
END_METHOD

END_INTERFACE

// Page/Page_PDEF/_Messages/_T_PDEF_Messages
(*
Description
===========
| Index: Array of messages on the PDEF page (see FB_Message)
| Method to clear message
*)
FUNCTION_BLOCK _T_PDEF_Messages IMPLEMENTS _I_T_PDEF_Messages_RO, _I_T_PDEF_Messages_Owner, _I_T_PDEF_Messages_Member, _I_T_PDEF_Messages_CopyFrom

VAR
	_Line		:	ARRAY[1..GVL_CONSTANT.MAX_PDEF_MESSAGES] OF _T_Message;	//ARRAY[1..GVL_CONSTANT.MAX_PDEF_MESSAGES] OF FB_Message
	_Dummy	:	_T_Message;
END_VAR

METHOD PUBLIC clear


VAR
	_index: INT;	//INT
END_VAR


FOR _index:= 1 TO GVL_CONSTANT.MAX_PDEF_MESSAGES DO
	_Line[_index].clear();
END_FOR
END_METHOD

METHOD PUBLIC CopyFrom
VAR_INPUT
	IN	: _I_T_PDEF_Messages_RO;
END_VAR

VAR
	_i: INT;
END_VAR

IF IN = 0 THEN RETURN;	END_IF

FOR _i:= 1 TO GVL_CONSTANT.MAX_PDEF_MESSAGES DO
	_Line[_i].CopyFrom(IN.Message_RO(_i));
END_FOR
END_METHOD

METHOD PUBLIC CopyTo
VAR_INPUT
	IN	: _I_T_PDEF_Messages_CopyFrom;
END_VAR

IF IN = 0 THEN RETURN;	END_IF

IN.CopyFrom(THIS^);
END_METHOD

METHOD PUBLIC Message : _I_T_Message
VAR_INPUT
	Number	: INT;
END_VAR

IF (Number < 1) OR (Number > GVL_CONSTANT.MAX_PDEF_MESSAGES) THEN	Message:= _Dummy;	RETURN;	END_IF

Message:= _Line[Number];
END_METHOD

METHOD PUBLIC Message_Owner : _I_T_Message_Owner
VAR_INPUT
	Number	: INT;
END_VAR

IF (Number < 1) OR (Number > GVL_CONSTANT.MAX_PDEF_MESSAGES) THEN	Message_Owner:= _Dummy;	RETURN;	END_IF

Message_Owner:= _Line[Number];
END_METHOD

METHOD PUBLIC Message_RO : _I_T_Message_RO
VAR_INPUT
	Number	: INT;
END_VAR

IF (Number < 1) OR (Number > GVL_CONSTANT.MAX_PDEF_MESSAGES) THEN	Message_RO:= _Dummy;	RETURN;	END_IF

Message_RO:= _Line[Number];
END_METHOD

END_FUNCTION_BLOCK

// Page/Page_PDEF/PDEF/FB_Page_PDEF
(*
:Author: Frank Dümpelmann <f.duempelmann@kostal.com>, Martin Hundt <m.hundt@kostal.com>
:Date: 2018-11-20

Function
========
Data structure representing the PDEF page of the user interface

Methods and Properties
======================
| Activate: Activate the Form
| Name: user defined Name of this page
| Message: Message Line under the Buttons (see FB_Message)
| Confirm: Big button at the bottom of PDEF Page
| Buttons: see FB_PDEF_Buttons
| Messages: Message Lines behind the Buttons (see FB_LISTING_Messages)
| Clear: Clear page
*)
FUNCTION_BLOCK PUBLIC FB_Page_PDEF IMPLEMENTS I_Page_PDEF_RO, I_Page_PDEF_Owner, I_Page_PDEF

VAR
	_Activate		: BOOL;	//BOOL	-	Activate the Form

	_Name			: KOSTAL_AF2024_Core_Settings.T_MaxString;	//Show a user defined Name of this page
	_Message	:	_T_Message;			//FB_Message - Message Line under the Buttons
	_Confirm	: _T_PDEF_Button;	//FB_PDEF_Button - Big button at the bottom of PDEF Page

	_Messages	:	_T_PDEF_Messages;	//FB_PDEF_Messages - Message Lines behind the Buttons

	_Buttons	: _T_PDEF_Buttons;	//FB_PDEF_Buttons
END_VAR

PROPERTY PUBLIC Buttons : _I_T_PDEF_Buttons_Member
GET

Buttons := _Buttons;
END_GET
END_PROPERTY

PROPERTY PUBLIC Confirm : _I_T_PDEF_Button_Member
GET

Confirm := _Confirm;
END_GET
END_PROPERTY

PROPERTY PUBLIC Message : _I_T_Message
GET

Message := _Message;
END_GET
END_PROPERTY

PROPERTY PUBLIC Messages : _I_T_PDEF_Messages_Member
GET

Messages := _Messages;
END_GET
END_PROPERTY

PROPERTY PUBLIC Buttons_Owner : _I_T_PDEF_Buttons_Owner
GET

Buttons_Owner := _Buttons;
END_GET
END_PROPERTY

PROPERTY PUBLIC Confirm_Owner : _I_T_PDEF_Button_Owner
GET

Confirm_Owner := _Confirm;
END_GET
END_PROPERTY

PROPERTY PUBLIC Message_Owner : _I_T_Message_Owner
GET

Message_Owner := _Message;
END_GET
END_PROPERTY

PROPERTY PUBLIC Messages_Owner : _I_T_PDEF_Messages_Owner
GET

Messages_Owner := _Messages;
END_GET
END_PROPERTY

PROPERTY PUBLIC Buttons_RO : _I_T_PDEF_Buttons_RO
GET

Buttons_RO := _Buttons;
END_GET
END_PROPERTY

PROPERTY PUBLIC Confirm_RO : _I_T_PDEF_Button_RO
GET

Confirm_RO := _Confirm;
END_GET
END_PROPERTY

PROPERTY PUBLIC Message_RO : _I_T_Message_RO
GET

Message_RO := _Message;
END_GET
END_PROPERTY

PROPERTY PUBLIC Messages_RO : _I_T_PDEF_Messages_RO
GET

Messages_RO := _Messages;
END_GET
END_PROPERTY

PROPERTY PUBLIC Activate : BOOL
GET


Activate:= _Activate;
END_GET
SET

_Activate:= Activate;
END_SET
END_PROPERTY

METHOD clear


_Activate		:= FALSE;

_Name	:= "";
_Message.clear();
_Confirm.clear();

_Buttons.clear();
_Messages.clear();
END_METHOD

PROPERTY PUBLIC Name : KOSTAL_AF2024_Core_Settings.T_MaxString
GET

Name:= _Name;
END_GET
SET

_Name:= Name;
END_SET
END_PROPERTY

END_FUNCTION_BLOCK

// Page/Page_PDEF/PDEF/I_Page_PDEF_RO
INTERFACE I_Page_PDEF_RO EXTENDS KOSTAL_AF2024_Core_System.I_Interface

PROPERTY PUBLIC Activate : BOOL
GET
END_GET
END_PROPERTY

PROPERTY PUBLIC Buttons_RO : _I_T_PDEF_Buttons_RO
GET
END_GET
END_PROPERTY

PROPERTY PUBLIC Confirm_RO : _I_T_PDEF_Button_RO
GET
END_GET
END_PROPERTY

PROPERTY PUBLIC Message_RO : _I_T_Message_RO
GET
END_GET
END_PROPERTY

PROPERTY PUBLIC Messages_RO : _I_T_PDEF_Messages_RO
GET
END_GET
END_PROPERTY

PROPERTY PUBLIC Name : KOSTAL_AF2024_Core_Settings.T_MaxString
GET
END_GET
END_PROPERTY

END_INTERFACE

// Page/Page_PDEF/PDEF/I_Page_PDEF_Owner
INTERFACE I_Page_PDEF_Owner EXTENDS I_Page_PDEF

PROPERTY PUBLIC Buttons : _I_T_PDEF_Buttons_Member
GET
END_GET
END_PROPERTY

PROPERTY PUBLIC Confirm : _I_T_PDEF_Button_Member
GET
END_GET
END_PROPERTY

PROPERTY PUBLIC Message : _I_T_Message
GET
END_GET
END_PROPERTY

PROPERTY PUBLIC Messages : _I_T_PDEF_Messages_Member
GET
END_GET
END_PROPERTY

PROPERTY PUBLIC Buttons_Owner : _I_T_PDEF_Buttons_Owner
GET
END_GET
END_PROPERTY

PROPERTY PUBLIC Confirm_Owner : _I_T_PDEF_Button_Owner
GET
END_GET
END_PROPERTY

PROPERTY PUBLIC Message_Owner : _I_T_Message_Owner
GET
END_GET
END_PROPERTY

PROPERTY PUBLIC Messages_Owner : _I_T_PDEF_Messages_Owner
GET
END_GET
END_PROPERTY

PROPERTY PUBLIC Buttons_RO : _I_T_PDEF_Buttons_RO
GET
END_GET
END_PROPERTY

PROPERTY PUBLIC Confirm_RO : _I_T_PDEF_Button_RO
GET
END_GET
END_PROPERTY

PROPERTY PUBLIC Message_RO : _I_T_Message_RO
GET
END_GET
END_PROPERTY

PROPERTY PUBLIC Messages_RO : _I_T_PDEF_Messages_RO
GET
END_GET
END_PROPERTY

PROPERTY PUBLIC Activate : BOOL
GET
END_GET
SET
END_SET
END_PROPERTY

METHOD clear
END_METHOD

PROPERTY PUBLIC Name : KOSTAL_AF2024_Core_Settings.T_MaxString
GET
END_GET
SET
END_SET
END_PROPERTY

END_INTERFACE

// Page/Page_PDEF/PDEF/I_Page_PDEF
INTERFACE I_Page_PDEF EXTENDS I_Page_PDEF_RO

PROPERTY PUBLIC Buttons : _I_T_PDEF_Buttons_Member
GET
END_GET
END_PROPERTY

PROPERTY PUBLIC Confirm : _I_T_PDEF_Button_Member
GET
END_GET
END_PROPERTY

PROPERTY PUBLIC Message : _I_T_Message
GET
END_GET
END_PROPERTY

PROPERTY PUBLIC Messages : _I_T_PDEF_Messages_Member
GET
END_GET
END_PROPERTY

PROPERTY PUBLIC Buttons_RO : _I_T_PDEF_Buttons_RO
GET
END_GET
END_PROPERTY

PROPERTY PUBLIC Confirm_RO : _I_T_PDEF_Button_RO
GET
END_GET
END_PROPERTY

PROPERTY PUBLIC Message_RO : _I_T_Message_RO
GET
END_GET
END_PROPERTY

PROPERTY PUBLIC Messages_RO : _I_T_PDEF_Messages_RO
GET
END_GET
END_PROPERTY

PROPERTY PUBLIC Activate : BOOL
GET
END_GET
SET
END_SET
END_PROPERTY

PROPERTY PUBLIC Name : KOSTAL_AF2024_Core_Settings.T_MaxString
GET
END_GET
SET
END_SET
END_PROPERTY

END_INTERFACE

// Page/Page_Station/FB_Page_Station
(*
:Author: Frank Dümpelmann <f.duempelmann@kostal.com>, Martin Hundt <m.hundt@kostal.com>
:Date: 2018-11-20

Function
========
Data structure representing the station page of the user interface

Methods and Properties
======================
| Activate: Activate the Form
| Deactivate: Deactivate the Form
| IsActiv: Response the state of the Form
| Buttons: see FB_LISTING_Buttons
| Messages: see FB_LISTING_Messages
*)
FUNCTION_BLOCK FB_Page_Station IMPLEMENTS I_Page_Station_RO, I_Page_Station_Owner, I_Page_Station

VAR
	_name	: KOSTAL_AF2024_Core_Settings.T_MaxString;

	_text	: KOSTAL_AF2024_Core_process.T_messageText_3_lines;	//KOSTAL_AF2024_Core_process.FB_messageText_3_lines
	_OnOff	: KOSTAL_AF2024_HMI_Controls.T_Button_controlled;	//KOSTAL_TC3_Controls_button.FB_Button_controlled
	_Minus	: KOSTAL_AF2024_HMI_Controls.T_Button_controlled;	//KOSTAL_TC3_Controls_button.FB_Button_controlled
	_Enter	: KOSTAL_AF2024_HMI_Controls.T_Button_controlled;	//KOSTAL_TC3_Controls_button.FB_Button_controlled
	_Plus	: KOSTAL_AF2024_HMI_Controls.T_Button_controlled;	//KOSTAL_TC3_Controls_button.FB_Button_controlled
	_Escape	: KOSTAL_AF2024_HMI_Controls.T_Button_controlled;	//KOSTAL_TC3_Controls_button.FB_Button_controlled
	
	_Custom	: _T_Fn_Button;

	_Status	: KOSTAL_AF2024_Core_process.FB_processCondition;	//KOSTAL_AF2024_Core_process.FB_processCondition
END_VAR

(*
Description
===========
| Enter button
*)
PROPERTY PUBLIC Button_Enter : KOSTAL_AF2024_HMI_Controls.I_T_Button_controlled
GET

Button_Enter := _Enter;
END_GET
END_PROPERTY

(*
Description
===========
| Escape button
*)
PROPERTY PUBLIC Button_Escape : KOSTAL_AF2024_HMI_Controls.I_T_Button_controlled
GET

Button_Escape := _Escape;
END_GET
END_PROPERTY

(*
Description
===========
| Minus/step back button
*)PROPERTY PUBLIC Button_Minus : KOSTAL_AF2024_HMI_Controls.I_T_Button_controlled
GET

Button_Minus := _Minus;
END_GET
END_PROPERTY

(*
Description
===========
| On/off button
*)
PROPERTY PUBLIC Button_OnOff : KOSTAL_AF2024_HMI_Controls.I_T_Button_controlled
GET

Button_OnOff := _OnOff;
END_GET
END_PROPERTY

(*
Description
===========
| Plus/step forward button
*)
PROPERTY PUBLIC Button_Plus : KOSTAL_AF2024_HMI_Controls.I_T_Button_controlled
GET

Button_Plus := _Plus;
END_GET
END_PROPERTY

(*
Description
===========
| Array of custom button
*)
PROPERTY PUBLIC Buttons_Custom : _I_T_Fn_Button
GET

Buttons_Custom := _Custom;
END_GET
END_PROPERTY

METHOD PUBLIC clear_controls

	
	_OnOff.clear_control();
	_Minus.clear_control();
	_Enter.clear_control();
	_Plus.clear_control();
	_Escape.clear_control();
	
	_Custom.clear_controls();
END_METHOD

PROPERTY PUBLIC Name : KOSTAL_AF2024_Core_Settings.T_MaxString
GET
Name := _name;
END_GET
SET
PUBLIC 
VAR
END_VAR
_name := Name;
END_SET
END_PROPERTY

(*
Description
===========
| Process condition of the station page (see FB_processCondition)
*)
PROPERTY PUBLIC Status : KOSTAL_AF2024_Core_process.I_processCondition_Owner
GET

Status := _Status;
END_GET
END_PROPERTY

(*
Description
===========
| Three lines of text to be displayed on the station page
*)
PROPERTY PUBLIC Text : KOSTAL_AF2024_Core_process.I_T_messageText_3_lines_Owner
GET

Text := _text;
END_GET
END_PROPERTY

(*
Description
===========
| Enter button
*)
PROPERTY PUBLIC Button_Enter_Owner : KOSTAL_AF2024_HMI_Controls.I_T_Button_controlled_Owner
GET

Button_Enter_Owner := _Enter;
END_GET
END_PROPERTY

(*
Description
===========
| Escape button
*)
PROPERTY PUBLIC Button_Escape_Owner : KOSTAL_AF2024_HMI_Controls.I_T_Button_controlled_Owner
GET

Button_Escape_Owner := _Escape;
END_GET
END_PROPERTY

(*
Description
===========
| Minus/step back button
*)PROPERTY PUBLIC Button_Minus_Owner : KOSTAL_AF2024_HMI_Controls.I_T_Button_controlled_Owner
GET

Button_Minus_Owner := _Minus;
END_GET
END_PROPERTY

(*
Description
===========
| On/off button
*)
PROPERTY PUBLIC Button_OnOff_Owner : KOSTAL_AF2024_HMI_Controls.I_T_Button_controlled_Owner
GET

Button_OnOff_Owner := _OnOff;
END_GET
END_PROPERTY

(*
Description
===========
| Plus/step forward button
*)
PROPERTY PUBLIC Button_Plus_Owner : KOSTAL_AF2024_HMI_Controls.I_T_Button_controlled_Owner
GET

Button_Plus_Owner := _Plus;
END_GET
END_PROPERTY

(*
Description
===========
| Array of custom button
*)
PROPERTY PUBLIC Buttons_Custom_Owner : _I_T_Fn_Button_Owner
GET

Buttons_Custom_Owner := _Custom;
END_GET
END_PROPERTY

METHOD PUBLIC clear

	_text.clear();

	_OnOff.clear();
	_Minus.clear();
	_Enter.clear();
	_Plus.clear();
	_Escape.clear();
	
	_Custom.clear();
	
	_Status.clear();

	_name:= "";
END_METHOD

METHOD PUBLIC clear_button

	
	_OnOff.clear();
	_Minus.clear();
	_Enter.clear();
	_Plus.clear();
	_Escape.clear();
	
	_Custom.clear();
END_METHOD

METHOD PUBLIC clear_signals

	
	_OnOff.clear_signals();
	_Minus.clear_signals();
	_Enter.clear_signals();
	_Plus.clear_signals();
	_Escape.clear_signals();
	
	_Custom.clear_signals();
END_METHOD

(*
Description
===========
| Process condition of the station page (see FB_processCondition)
*)
PROPERTY PUBLIC Status_Owner : KOSTAL_AF2024_Core_process.I_processCondition_Owner
GET

Status_Owner := _Status;
END_GET
END_PROPERTY

(*
Description
===========
| Three lines of text to be displayed on the station page
*)
PROPERTY PUBLIC Text_Owner : KOSTAL_AF2024_Core_process.I_T_messageText_3_lines_Owner
GET

Text_Owner := _text;
END_GET
END_PROPERTY

(*
Description
===========
| Enter button
*)
PROPERTY PUBLIC Button_Enter_RO : KOSTAL_AF2024_HMI_Controls.I_T_Button_controlled
GET

Button_Enter_RO := _Enter;
END_GET
END_PROPERTY

(*
Description
===========
| Escape button
*)
PROPERTY PUBLIC Button_Escape_RO : I_T_Button_controlled
GET

Button_Escape_RO := _Escape;
END_GET
END_PROPERTY

(*
Description
===========
| Minus/step back button
*)PROPERTY PUBLIC Button_Minus_RO : I_T_Button_controlled
GET

Button_Minus_RO := _Minus;
END_GET
END_PROPERTY

(*
Description
===========
| On/off button
*)
PROPERTY PUBLIC Button_OnOff_RO : I_T_Button_controlled
GET

Button_OnOff_RO := _OnOff;
END_GET
END_PROPERTY

(*
Description
===========
| Plus/step forward button
*)
PROPERTY PUBLIC Button_Plus_RO : I_T_Button_controlled
GET

Button_Plus_RO := _Plus;
END_GET
END_PROPERTY

(*
Description
===========
| Array of custom button
*)
PROPERTY PUBLIC Buttons_Custom_RO : _I_T_Fn_Button_RO
GET

Buttons_Custom_RO := _Custom;
END_GET
END_PROPERTY

PROPERTY PUBLIC Name_RO : KOSTAL_AF2024_Core_Settings.T_MaxString
GET
Name_RO := _name;
END_GET
END_PROPERTY

(*
Description
===========
| Process condition of the station page (see FB_processCondition)
*)
PROPERTY PUBLIC Status_RO : KOSTAL_AF2024_Core_Process.I_processCondition
GET

Status_RO := _Status;
END_GET
END_PROPERTY

(*
Description
===========
| Three lines of text to be displayed on the station page
*)
PROPERTY PUBLIC Text_RO : KOSTAL_AF2024_Core_process.I_T_messageText_3_lines
GET

Text_RO := _text;
END_GET
END_PROPERTY

END_FUNCTION_BLOCK

// Page/Page_Station/I_Page_Station_RO
INTERFACE I_Page_Station_RO EXTENDS KOSTAL_AF2024_Core_System.I_Interface

(*
Description
===========
| Enter button
*)
PROPERTY PUBLIC Button_Enter_RO : KOSTAL_AF2024_HMI_Controls.I_T_Button_controlled
GET
END_GET
END_PROPERTY

(*
Description
===========
| Escape button
*)
PROPERTY PUBLIC Button_Escape_RO : KOSTAL_AF2024_HMI_Controls.I_T_Button_controlled
GET
END_GET
END_PROPERTY

(*
Description
===========
| Minus/step back button
*)PROPERTY PUBLIC Button_Minus_RO : KOSTAL_AF2024_HMI_Controls.I_T_Button_controlled
GET
END_GET
END_PROPERTY

(*
Description
===========
| On/off button
*)
PROPERTY PUBLIC Button_OnOff_RO : KOSTAL_AF2024_HMI_Controls.I_T_Button_controlled
GET
END_GET
END_PROPERTY

(*
Description
===========
| Plus/step forward button
*)
PROPERTY PUBLIC Button_Plus_RO : KOSTAL_AF2024_HMI_Controls.I_T_Button_controlled
GET
END_GET
END_PROPERTY

(*
Description
===========
| Array of custom button
*)
PROPERTY PUBLIC Buttons_Custom_RO : _I_T_Fn_Button_RO
GET
END_GET
END_PROPERTY

PROPERTY PUBLIC Name : KOSTAL_AF2024_Core_Settings.T_MaxString
GET
END_GET
END_PROPERTY

(*
Description
===========
| Process condition of the station page (see FB_processCondition)
*)
PROPERTY PUBLIC Status_RO : KOSTAL_AF2024_Core_process.I_processCondition
GET
END_GET
END_PROPERTY

(*
Description
===========
| Three lines of text to be displayed on the station page
*)
PROPERTY PUBLIC Text_RO : KOSTAL_AF2024_Core_process.I_T_messageText_3_lines
GET
END_GET
END_PROPERTY

END_INTERFACE

// Page/Page_Station/I_Page_Station_Owner
INTERFACE I_Page_Station_Owner EXTENDS I_Page_Station

(*
Description
===========
| Enter button
*)
PROPERTY PUBLIC Button_Enter_Owner : I_T_Button_controlled_Owner
GET
END_GET
END_PROPERTY

(*
Description
===========
| Escape button
*)
PROPERTY PUBLIC Button_Escape_Owner : I_T_Button_controlled_Owner
GET
END_GET
END_PROPERTY

(*
Description
===========
| Minus/step back button
*)PROPERTY PUBLIC Button_Minus_Owner : I_T_Button_controlled_Owner
GET
END_GET
END_PROPERTY

(*
Description
===========
| On/off button
*)
PROPERTY PUBLIC Button_OnOff_Owner : I_T_Button_controlled_Owner
GET
END_GET
END_PROPERTY

(*
Description
===========
| Plus/step forward button
*)
PROPERTY PUBLIC Button_Plus_Owner : I_T_Button_controlled_Owner
GET
END_GET
END_PROPERTY

(*
Description
===========
| Array of custom button
*)
PROPERTY PUBLIC Buttons_Custom_Owner : _I_T_Fn_Button_Owner
GET
END_GET
END_PROPERTY

METHOD PUBLIC clear
END_METHOD

METHOD PUBLIC clear_button
END_METHOD

METHOD PUBLIC clear_signals
END_METHOD

(*
Description
===========
| Process condition of the station page (see FB_processCondition)
*)
PROPERTY PUBLIC Status_Owner : KOSTAL_AF2024_Core_process.I_processCondition_Owner
GET
END_GET
END_PROPERTY

(*
Description
===========
| Three lines of text to be displayed on the station page
*)
PROPERTY PUBLIC Text_Owner : KOSTAL_AF2024_Core_process.I_T_messageText_3_lines_Owner
GET
END_GET
END_PROPERTY

END_INTERFACE

// Page/Page_Station/I_Page_Station
INTERFACE I_Page_Station EXTENDS I_Page_Station_RO

(*
Description
===========
| Enter button
*)
PROPERTY PUBLIC Button_Enter : KOSTAL_AF2024_HMI_Controls.I_T_Button_controlled
GET
END_GET
END_PROPERTY

(*
Description
===========
| Escape button
*)
PROPERTY PUBLIC Button_Escape : KOSTAL_AF2024_HMI_Controls.I_T_Button_controlled
GET
END_GET
END_PROPERTY

(*
Description
===========
| Minus/step back button
*)PROPERTY PUBLIC Button_Minus : KOSTAL_AF2024_HMI_Controls.I_T_Button_controlled
GET
END_GET
END_PROPERTY

(*
Description
===========
| On/off button
*)
PROPERTY PUBLIC Button_OnOff : KOSTAL_AF2024_HMI_Controls.I_T_Button_controlled
GET
END_GET
END_PROPERTY

(*
Description
===========
| Plus/step forward button
*)
PROPERTY PUBLIC Button_Plus : KOSTAL_AF2024_HMI_Controls.I_T_Button_controlled
GET
END_GET
END_PROPERTY

(*
Description
===========
| Array of custom button
*)
PROPERTY PUBLIC Buttons_Custom : _I_T_Fn_Button
GET
END_GET
END_PROPERTY

METHOD PUBLIC clear_controls
END_METHOD

PROPERTY PUBLIC Name : KOSTAL_AF2024_Core_Settings.T_MaxString
SET
END_SET
END_PROPERTY

(*
Description
===========
| Process condition of the station page (see FB_processCondition)
*)
PROPERTY PUBLIC Status : KOSTAL_AF2024_Core_process.I_processCondition_Owner
GET
END_GET
END_PROPERTY

(*
Description
===========
| Three lines of text to be displayed on the station page
*)
PROPERTY PUBLIC Text : KOSTAL_AF2024_Core_process.I_T_messageText_3_lines_Owner
GET
END_GET
END_PROPERTY

END_INTERFACE

// Page/Page_XYZ/_Buttons/_I_T_XYZ_Buttons
INTERFACE _I_T_XYZ_Buttons EXTENDS _I_T_XYZ_Buttons_RO

METHOD PUBLIC Button : KOSTAL_AF2024_HMI_Controls.I_T_Button_controlled
VAR_INPUT
	Number	: INT;
END_VAR
END_METHOD

METHOD PUBLIC clear_controls
END_METHOD

END_INTERFACE

// Page/Page_XYZ/_Buttons/_I_T_XYZ_Buttons_RO
INTERFACE _I_T_XYZ_Buttons_RO EXTENDS KOSTAL_AF2024_Core_System.I_Interface

METHOD PUBLIC Button_RO : KOSTAL_AF2024_HMI_Controls.I_T_Button_controlled_RO
VAR_INPUT
	Number	: INT;
END_VAR
END_METHOD

METHOD PUBLIC CopyTo
VAR_INPUT
END_VAR
END_METHOD

END_INTERFACE

// Page/Page_XYZ/_Buttons/_I_T_XYZ_Buttons_CopyFrom
INTERFACE _I_T_XYZ_Buttons_CopyFrom EXTENDS KOSTAL_AF2024_Core_System.I_Interface

METHOD PUBLIC CopyFrom
VAR_INPUT
	IN	: _I_T_Listing_Buttons_RO;
END_VAR
END_METHOD

END_INTERFACE

// Page/Page_XYZ/_Buttons/_I_T_XYZ_Buttons_Owner
INTERFACE _I_T_XYZ_Buttons_Owner EXTENDS _I_T_XYZ_Buttons

METHOD PUBLIC Button_Owner : KOSTAL_AF2024_HMI_Controls.I_T_Button_controlled_Owner
VAR_INPUT
	Number	: INT;
END_VAR
END_METHOD

METHOD PUBLIC clear
END_METHOD

METHOD PUBLIC clear_signals
END_METHOD

METHOD PUBLIC CopyFrom
VAR_INPUT
	IN	: _I_T_Listing_Buttons_RO;
END_VAR
END_METHOD

END_INTERFACE

// Page/Page_XYZ/_Buttons/_T_XYZ_Buttons
(*

:Author: Frank Dümpelmann <f.duempelmann@kostal.com>, Martin Hundt <m.hundt@kostal.com>
:Date: 2018-11-20

Function
========
Data structure representing the custom buttons in the XYZ page of the user interface

Methods and Properties
======================
| _customButtons: Array with Buttons (see FB_Button_controlled)
| clear signals of buttons
| clear all buttons
*)
FUNCTION_BLOCK _T_XYZ_Buttons IMPLEMENTS _I_T_XYZ_Buttons_RO, _I_T_XYZ_Buttons_Owner, _I_T_XYZ_Buttons, _I_T_XYZ_Buttons_CopyFrom

VAR
	_customButtons	: ARRAY[1..GVL_CONSTANT.MAX_XYZ_BUTTON] OF KOSTAL_AF2024_HMI_Controls.T_Button_controlled;
	
	_Dummy	: KOSTAL_AF2024_HMI_Controls.T_Button_controlled;
END_VAR

METHOD PUBLIC Button : KOSTAL_AF2024_HMI_Controls.I_T_Button_controlled
VAR_INPUT
	Number	: INT;
END_VAR
IF (Number < 1) OR (Number > GVL_CONSTANT.MAX_XYZ_BUTTON) THEN	
	Button:= _Dummy;	
	RETURN;	
END_IF

	
Button:= _customButtons[Number];
END_METHOD

METHOD PUBLIC Button_Owner : KOSTAL_AF2024_HMI_Controls.I_T_Button_controlled_Owner
VAR_INPUT
	Number	: INT;
END_VAR

IF (Number < 1) OR (Number > GVL_CONSTANT.MAX_XYZ_BUTTON) THEN	
	Button_Owner:= _Dummy;	
	RETURN;	
END_IF

	
Button_Owner:= _customButtons[Number];
END_METHOD

METHOD PUBLIC Button_RO : KOSTAL_AF2024_HMI_Controls.I_T_Button_controlled_RO
VAR_INPUT
	Number	: INT;
END_VAR

IF (Number < 1) OR (Number > GVL_CONSTANT.MAX_XYZ_BUTTON) THEN	
	Button_RO:= _Dummy;	
	RETURN;	
END_IF

	
Button_RO:= _customButtons[Number];
END_METHOD

METHOD PUBLIC clear


VAR
	_index: INT;	//INT
END_VAR


FOR _index:= 1 TO GVL_CONSTANT.MAX_XYZ_BUTTON DO
	_customButtons[_index].clear();
END_FOR
END_METHOD

METHOD PUBLIC clear_controls


VAR
	_index: INT;	//INT
END_VAR


FOR _index:= 1 TO GVL_CONSTANT.MAX_XYZ_BUTTON DO
	_customButtons[_index].clear_control();
END_FOR
END_METHOD

METHOD PUBLIC clear_signals


VAR
	_index: INT;	//INT
END_VAR


FOR _index:= 1 TO GVL_CONSTANT.MAX_XYZ_BUTTON DO
	_customButtons[_index].clear_signals();
END_FOR
END_METHOD

METHOD PUBLIC CopyFrom
VAR_INPUT
	IN	: _I_T_Listing_Buttons_RO;
END_VAR

VAR
	_i: INT;
END_VAR

IF IN = 0 THEN RETURN;	END_IF

FOR _i:= 1 TO GVL_CONSTANT.MAX_XYZ_BUTTON DO
	_customButtons[_i].CopyFrom(IN.Button_RO(_i));
END_FOR
END_METHOD

METHOD PUBLIC CopyTo
VAR_INPUT
END_VAR
END_METHOD

END_FUNCTION_BLOCK

// Page/Page_XYZ/FB_page_XYZ
(*

:Author: Frank Dümpelmann <f.duempelmann@kostal.com>, Martin Hundt <m.hundt@kostal.com>
:Date: 2020-02-28

Function
========
Data structure representing the XYZ page in the user Interface

Methods and Properties
======================
| activate: Page is activated
| text: Four lines of text in the page
| clear all or signals only
| other properties represent the buttons on the page
*)
FUNCTION_BLOCK PUBLIC FB_page_XYZ IMPLEMENTS I_page_XYZ_RO, I_page_XYZ_Owner, I_page_XYZ

VAR
		_text	:	ARRAY [1..4] OF KOSTAL_AF2024_Core_Settings.T_MaxString;
		
		_Activate	: BOOL;	//BOOL	-	Activate the Form
		_IsActiv	: BOOL;	//BOOL	-	Response the state of the Form

		_Forward	: KOSTAL_AF2024_HMI_Controls.T_Button_controlled;	//KOSTAL_TC3_Controls_button.FB_Button_controlled
		_Backward	: KOSTAL_AF2024_HMI_Controls.T_Button_controlled;	//KOSTAL_TC3_Controls_button.FB_Button_controlled
		_Right		: KOSTAL_AF2024_HMI_Controls.T_Button_controlled;	//KOSTAL_TC3_Controls_button.FB_Button_controlled
		_Left		: KOSTAL_AF2024_HMI_Controls.T_Button_controlled;	//KOSTAL_TC3_Controls_button.FB_Button_controlled
		_Up			: KOSTAL_AF2024_HMI_Controls.T_Button_controlled;	//KOSTAL_TC3_Controls_button.FB_Button_controlled
		_Down		: KOSTAL_AF2024_HMI_Controls.T_Button_controlled;	//KOSTAL_TC3_Controls_button.FB_Button_controlled
		


		_Plus		: KOSTAL_AF2024_HMI_Controls.T_Button_controlled;	//KOSTAL_TC3_Controls_button.FB_Button_controlled
		_Minus		: KOSTAL_AF2024_HMI_Controls.T_Button_controlled;	//KOSTAL_TC3_Controls_button.FB_Button_controlled
		
		_Custom	: _T_XYZ_Buttons;
END_VAR

PROPERTY PUBLIC Button_Backward : KOSTAL_AF2024_HMI_Controls.I_T_Button_controlled
GET

Button_Backward := _Backward;
END_GET
END_PROPERTY

PROPERTY PUBLIC Button_Down : KOSTAL_AF2024_HMI_Controls.I_T_Button_controlled
GET

Button_Down := _Down;
END_GET
END_PROPERTY

PROPERTY PUBLIC Button_Forward : KOSTAL_AF2024_HMI_Controls.I_T_Button_controlled
GET

Button_Forward := _Forward;
END_GET
END_PROPERTY

PROPERTY PUBLIC Button_Left : KOSTAL_AF2024_HMI_Controls.I_T_Button_controlled
GET

Button_Left := _Left;
END_GET
END_PROPERTY

PROPERTY PUBLIC Button_Minus : KOSTAL_AF2024_HMI_Controls.I_T_Button_controlled
GET

Button_Minus := _Minus;
END_GET
END_PROPERTY

PROPERTY PUBLIC Button_Plus : KOSTAL_AF2024_HMI_Controls.I_T_Button_controlled
GET

Button_Plus := _Plus;
END_GET
END_PROPERTY

PROPERTY PUBLIC Button_Right : KOSTAL_AF2024_HMI_Controls.I_T_Button_controlled
GET

Button_Right := _Right;
END_GET
END_PROPERTY

PROPERTY PUBLIC Button_Up : KOSTAL_AF2024_HMI_Controls.I_T_Button_controlled
GET

Button_Up := _Up;
END_GET
END_PROPERTY

(*
Description
===========
| Array of custom button
*)
PROPERTY PUBLIC Buttons_Custom : _I_T_XYZ_Buttons
GET

Buttons_Custom := _Custom;
END_GET
END_PROPERTY

{}
METHOD PUBLIC clear_controls



_Forward.clear_control();
_Backward.clear_control();
_Down.clear_control();
_Left.clear_control();
_Minus.clear_control();
_Plus.clear_control();
_Right.clear_control();
_Up.clear_control();
END_METHOD

METHOD PUBLIC SetText : BOOL
VAR_INPUT
	Line	: USINT;
	Text	: KOSTAL_AF2024_Core_Settings.T_MaxString;	
END_VAR
IF (Line < 1) OR (Line > GVL_CONSTANT.MAX_XYZ_LINE) THEN	RETURN;	END_IF

_text[Line]:= Text;

SetText:= TRUE;
END_METHOD

PROPERTY PUBLIC Button_Backward_Owner : KOSTAL_AF2024_HMI_Controls.I_T_Button_controlled_Owner
GET

Button_Backward_Owner := _Backward;
END_GET
END_PROPERTY

PROPERTY PUBLIC Button_Down_Owner : KOSTAL_AF2024_HMI_Controls.I_T_Button_controlled_Owner
GET

Button_Down_Owner := _Down;
END_GET
END_PROPERTY

PROPERTY PUBLIC Button_Forward_Owner : KOSTAL_AF2024_HMI_Controls.I_T_Button_controlled_Owner
GET

Button_Forward_Owner := _Forward;
END_GET
END_PROPERTY

PROPERTY PUBLIC Button_Left_Owner : KOSTAL_AF2024_HMI_Controls.I_T_Button_controlled_Owner
GET

Button_Left_Owner := _Left;
END_GET
END_PROPERTY

PROPERTY PUBLIC Button_Minus_Owner : KOSTAL_AF2024_HMI_Controls.I_T_Button_controlled_Owner
GET

Button_Minus_Owner := _Minus;
END_GET
END_PROPERTY

PROPERTY PUBLIC Button_Plus_Owner : KOSTAL_AF2024_HMI_Controls.I_T_Button_controlled_Owner
GET

Button_Plus_Owner := _Plus;
END_GET
END_PROPERTY

PROPERTY PUBLIC Button_Right_Owner : KOSTAL_AF2024_HMI_Controls.I_T_Button_controlled_Owner
GET

Button_Right_Owner := _Right;
END_GET
END_PROPERTY

PROPERTY PUBLIC Button_Up_Owner : KOSTAL_AF2024_HMI_Controls.I_T_Button_controlled_Owner
GET

Button_Up_Owner := _Up;
END_GET
END_PROPERTY

(*
Description
===========
| Array of custom button
*)
PROPERTY PUBLIC Buttons_Custom_Owner : _I_T_XYZ_Buttons_Owner
GET

Buttons_Custom_Owner := _Custom;
END_GET
END_PROPERTY

PROPERTY PUBLIC Button_Backward_RO : KOSTAL_AF2024_HMI_Controls.I_T_Button_controlled
GET

Button_Backward_RO := _Backward;
END_GET
END_PROPERTY

PROPERTY PUBLIC Button_Down_RO : KOSTAL_AF2024_HMI_Controls.I_T_Button_controlled
GET

Button_Down_RO := _Down;
END_GET
END_PROPERTY

PROPERTY PUBLIC Button_Forward_RO : KOSTAL_AF2024_HMI_Controls.I_T_Button_controlled
GET

Button_Forward_RO := _Forward;
END_GET
END_PROPERTY

PROPERTY PUBLIC Button_Left_RO : KOSTAL_AF2024_HMI_Controls.I_T_Button_controlled
GET

Button_Left_RO := _Left;
END_GET
END_PROPERTY

PROPERTY PUBLIC Button_Minus_RO : KOSTAL_AF2024_HMI_Controls.I_T_Button_controlled
GET

Button_Minus_RO := _Minus;
END_GET
END_PROPERTY

PROPERTY PUBLIC Button_Plus_RO : KOSTAL_AF2024_HMI_Controls.I_T_Button_controlled
GET

Button_Plus_RO := _Plus;
END_GET
END_PROPERTY

PROPERTY PUBLIC Button_Right_RO : KOSTAL_AF2024_HMI_Controls.I_T_Button_controlled
GET

Button_Right_RO := _Right;
END_GET
END_PROPERTY

PROPERTY PUBLIC Button_Up_RO : KOSTAL_AF2024_HMI_Controls.I_T_Button_controlled
GET

Button_Up_RO := _Up;
END_GET
END_PROPERTY

(*
Description
===========
| Array of custom button
*)
PROPERTY PUBLIC Buttons_Custom_RO : _I_T_XYZ_Buttons_RO
GET

Buttons_Custom_RO := _Custom;
END_GET
END_PROPERTY

METHOD PUBLIC GetText : KOSTAL_AF2024_Core_Settings.T_MaxString
VAR_INPUT
	Line	: USINT;
END_VAR

IF (Line < 1) OR (Line > GVL_CONSTANT.MAX_XYZ_LINE) THEN	RETURN;	END_IF

GetText:= _Text[Line];
END_METHOD

PROPERTY PUBLIC Activate : BOOL
GET

Activate:= _Activate;
END_GET
SET

_Activate:= Activate;
END_SET
END_PROPERTY

//Clear hole content
METHOD PUBLIC clear


VAR
	_index: INT;	//INT
END_VAR


_Forward.clear();
_Backward.clear();
_Down.clear();
_Left.clear();
_Minus.clear();
_Plus.clear();
_Right.clear();
_Up.clear();

FOR _index:= 1 TO 4 DO
	_text[_index]:= "";
END_FOR
		
_Activate	:= FALSE;
_IsActiv	:= FALSE;
END_METHOD

{}
METHOD PUBLIC clear_signals


_Forward.clear_signals();
_Backward.clear_signals();
_Down.clear_signals();
_Left.clear_signals();
_Minus.clear_signals();
_Plus.clear_signals();
_Right.clear_signals();
_Up.clear_signals();
END_METHOD

END_FUNCTION_BLOCK

// Page/Page_XYZ/I_page_XYZ_RO
INTERFACE I_page_XYZ_RO EXTENDS KOSTAL_AF2024_Core_System.I_Interface

PROPERTY PUBLIC Activate : BOOL
GET
END_GET
END_PROPERTY

PROPERTY PUBLIC Button_Backward_RO : KOSTAL_AF2024_HMI_Controls.I_T_Button_controlled
GET
END_GET
END_PROPERTY

PROPERTY PUBLIC Button_Down_RO : KOSTAL_AF2024_HMI_Controls.I_T_Button_controlled
GET
END_GET
END_PROPERTY

PROPERTY PUBLIC Button_Forward_RO : KOSTAL_AF2024_HMI_Controls.I_T_Button_controlled
GET
END_GET
END_PROPERTY

PROPERTY PUBLIC Button_Left_RO : KOSTAL_AF2024_HMI_Controls.I_T_Button_controlled
GET
END_GET
END_PROPERTY

PROPERTY PUBLIC Button_Minus_RO : KOSTAL_AF2024_HMI_Controls.I_T_Button_controlled
GET
END_GET
END_PROPERTY

PROPERTY PUBLIC Button_Plus_RO : KOSTAL_AF2024_HMI_Controls.I_T_Button_controlled
GET
END_GET
END_PROPERTY

PROPERTY PUBLIC Button_Right_RO : KOSTAL_AF2024_HMI_Controls.I_T_Button_controlled
GET
END_GET
END_PROPERTY

PROPERTY PUBLIC Button_Up_RO : KOSTAL_AF2024_HMI_Controls.I_T_Button_controlled
GET
END_GET
END_PROPERTY

METHOD PUBLIC GetText : KOSTAL_AF2024_Core_Settings.T_MaxString
VAR_INPUT
	Line	: USINT;
END_VAR
END_METHOD

END_INTERFACE

// Page/Page_XYZ/I_page_XYZ_Owner
INTERFACE I_page_XYZ_Owner EXTENDS I_page_XYZ

PROPERTY PUBLIC Button_Backward_Owner : KOSTAL_AF2024_HMI_Controls.I_T_Button_controlled_Owner
GET
END_GET
END_PROPERTY

PROPERTY PUBLIC Button_Down_Owner : KOSTAL_AF2024_HMI_Controls.I_T_Button_controlled_Owner
GET
END_GET
END_PROPERTY

PROPERTY PUBLIC Button_Forward_Owner : KOSTAL_AF2024_HMI_Controls.I_T_Button_controlled_Owner
GET
END_GET
END_PROPERTY

PROPERTY PUBLIC Button_Left_Owner : KOSTAL_AF2024_HMI_Controls.I_T_Button_controlled_Owner
GET
END_GET
END_PROPERTY

PROPERTY PUBLIC Button_Minus_Owner : KOSTAL_AF2024_HMI_Controls.I_T_Button_controlled_Owner
GET
END_GET
END_PROPERTY

PROPERTY PUBLIC Button_Plus_Owner : KOSTAL_AF2024_HMI_Controls.I_T_Button_controlled_Owner
GET
END_GET
END_PROPERTY

PROPERTY PUBLIC Button_Right_Owner : KOSTAL_AF2024_HMI_Controls.I_T_Button_controlled_Owner
GET
END_GET
END_PROPERTY

PROPERTY PUBLIC Button_Up_Owner : KOSTAL_AF2024_HMI_Controls.I_T_Button_controlled_Owner
GET
END_GET
END_PROPERTY

//Clear hole content
METHOD PUBLIC clear
END_METHOD

{}
METHOD PUBLIC clear_signals
END_METHOD

END_INTERFACE

// Page/Page_XYZ/I_page_XYZ
INTERFACE I_page_XYZ EXTENDS I_page_XYZ_RO

PROPERTY PUBLIC Activate : BOOL
GET
END_GET
SET
END_SET
END_PROPERTY

PROPERTY PUBLIC Button_Backward : KOSTAL_AF2024_HMI_Controls.I_T_Button_controlled
GET
END_GET
END_PROPERTY

PROPERTY PUBLIC Button_Down : KOSTAL_AF2024_HMI_Controls.I_T_Button_controlled
GET
END_GET
END_PROPERTY

PROPERTY PUBLIC Button_Forward : KOSTAL_AF2024_HMI_Controls.I_T_Button_controlled
GET
END_GET
END_PROPERTY

PROPERTY PUBLIC Button_Left : KOSTAL_AF2024_HMI_Controls.I_T_Button_controlled
GET
END_GET
END_PROPERTY

PROPERTY PUBLIC Button_Minus : KOSTAL_AF2024_HMI_Controls.I_T_Button_controlled
GET
END_GET
END_PROPERTY

PROPERTY PUBLIC Button_Plus : KOSTAL_AF2024_HMI_Controls.I_T_Button_controlled
GET
END_GET
END_PROPERTY

PROPERTY PUBLIC Button_Right : KOSTAL_AF2024_HMI_Controls.I_T_Button_controlled
GET
END_GET
END_PROPERTY

PROPERTY PUBLIC Button_Up : KOSTAL_AF2024_HMI_Controls.I_T_Button_controlled
GET
END_GET
END_PROPERTY

{}
METHOD PUBLIC clear_controls
END_METHOD

METHOD PUBLIC SetText : BOOL
VAR_INPUT
	Line	: USINT;
	Text	: KOSTAL_AF2024_Core_Settings.T_MaxString;	
END_VAR
END_METHOD

END_INTERFACE

// Project Information/F_GetCompany
// This function has been automatically generated from the project information.
{attribute 'signature_flag' := '1073741824'}
{attribute 'TcGenerated'}
{attribute 'no-analysis'}
FUNCTION F_GetCompany : WSTRING
VAR_INPUT
	
END_VAR

F_GetCompany := "KOSTAL GmbH & Co.KG";

END_FUNCTION

// Project Information/F_GetTitle
// This function has been automatically generated from the project information.
{attribute 'signature_flag' := '1073741824'}
{attribute 'TcGenerated'}
{attribute 'no-analysis'}
FUNCTION F_GetTitle : WSTRING
VAR_INPUT
	
END_VAR

F_GetTitle := "KOSTAL.AF2024.HMI.I_Hmi";

END_FUNCTION

// Project Information/F_GetVersion
// This function has been automatically generated from the project information.
{attribute 'signature_flag' := '1073741824'}
{attribute 'TcGenerated'}
{attribute 'no-analysis'}
FUNCTION F_GetVersion : ST_LibVersion
VAR_INPUT
	
END_VAR

F_GetVersion.iMajor := 1;
F_GetVersion.iMinor := 0;
F_GetVersion.iBuild := 0;
F_GetVersion.iRevision := 0;
F_GetVersion.sVersion := '1.0.0.0';
F_GetVersion.nFlags := 0;

END_FUNCTION
